                           //Feedback
                           "Mode_HMI_Feedback_Tag(1)" := "Control_DB".LCnv_Control[#i].Mode;
                           "Enabled_HMI_Feedback_Tag(1)" := "Control_DB".LCnv_Control[#i].Enabled;
                           "Error_HMI_Feedback_Tag(1)" := "Control_DB".LCnv_Control[#i].Error;
                           "Warning_HMI_Feedback_Tag(1)" := "Control_DB".LCnv_Control[#i].Warning;
                           "Stopped_HMI_Feedback_Tag(1)" := "Control_DB".LCnv_Control[#i].Stopped;
                           "Running_HMI_Feedback_Tag(1)" := "Control_DB".LCnv_Control[#i].Running;
                           "Ready_For_Task_HMI_Feedback_Tag(1)" := "Control_DB".LCnv_Control[#i].Ready_For_Task;
                           "Cnv_Occupied_HMI_Feedback_Tag(1)" := "Control_DB".LCnv_Control[#i].Cnv_Occupied;
                           "Shuttle_in_place_HMI_Feedback_Tag(1)" := "Control_DB".LCnv_Control[#i].Shuttle_In_Place;
                           "Current_Task_Type_HMI_Feedback_Tag(1)" := "Control_DB".LCnv_Control[#i].Current_Task_Type;
                           "Current_Task_ID_HMI_Feedback_Tag(1)" := "Control_DB".LCnv_Control[#i].Current_Task_ID;
                           "SM_State_HMI_Feedback_Tag(1)" := "Control_DB".LCnv_Control[#i].SM_State;
                           IF "Control_DB".LCnv_Control[#i].Motor.Forward THEN
                               "Motor_Direction_HMI_Feedback_Tag(1)" := 1;
                           ELSIF "Control_DB".LCnv_Control[#i].Motor.Reverse THEN
                               "Motor_Direction_HMI_Feedback_Tag(1)" := 2;
                           ELSE
                               "Motor_Direction_HMI_Feedback_Tag(1)" := 0;
                           END_IF;
                           "Motor_Speed_Requested_HMI_Feedback_Tag(1)" := "Control_DB".LCnv_Control[#i].Motor.Speed;
                           "Motor_Speed_Actual_HMI_Feedback_Tag(1)" := "Control_DB".LCnv_Control[#i].Motor.Speed_Actual;
                           "Transfer_To_ID_HMI_Tag(1)" := "Control_DB".LCnv_Control[#i].Instruction.Transfer_To_ID;
                           "Transfer_From_ID_HMI_Tag(1)" := "Control_DB".LCnv_Control[#i].Instruction.Transfer_From_ID;

                           //Instructions
                           IF "HMI_DB".ScreenNo = 2 THEN
                               "Control_DB".LCnv_Control[#i].Instruction.Stop := "Stop_HMI_Tag(1)";
                               "Control_DB".LCnv_Control[#i].Instruction.Execute := "Manual_Fwd_HMI_Tag(1)" OR "Manual_Bwd_HMI_Tag(1)";
                               "Control_DB".LCnv_Control[#i].Instruction.Mode_Change := "Mode_Change_HMI_Tag(1)";
                               "Control_DB".LCnv_Control[#i].Instruction.Enable := "Enable_HMI_Tag(1)";
                               IF "Control_DB".LCnv_Control[#i].Mode <> 3 THEN
                                   "Control_DB".LCnv_Control[#i].Instruction.Foward := "Manual_Fwd_HMI_Tag(1)";
                                   "Control_DB".LCnv_Control[#i].Instruction.Backward := "Manual_Bwd_HMI_Tag(1)";
                                   "Control_DB".LCnv_Control[#i].Instruction.Start_Transfer := "Start_Transfer_HMI_Tag(1)";
                                   IF "Control_DB".LCnv_Control[#i].Mode = 1 THEN
                                       "Control_DB".LCnv_Control[#i].Instruction.Start_Transfer_Backward := "Transfer_Backward(1)";
                                   END_IF;
                                   "Control_DB".LCnv_Control[#i].Safety_Stop_Cnrl.Instruction.Manual_Extend := "Manual_Sfty_Stopper_Up(1)";
                                   "Control_DB".LCnv_Control[#i].Safety_Stop_Cnrl.Instruction.Manual_Retract := "Manual_Sfty_Stopper_Down(1)";

                                   "Control_DB".LCnv_Control[#i].Instruction.Task_ID := "Task_ID_HMI_Tag(1)";
                                   // "Control_DB".LCnv_Control[#i].Instruction.Transfer_To_ID := "Transfer_To_ID_HMI_Tag(1)";
                                   // "Control_DB".LCnv_Control[#i].Instruction.Transfer_From_ID := "Transfer_From_ID_HMI_Tag(1)";
                                   IF "CNV_In_Out(1)" THEN // 0 = Inbound, 1 = Outbound
                                       "Control_DB".LCnv_Control[#i].Instruction.Transfer_To_ID := DINT#120001 + (#i * 100);
                                       "Control_DB".LCnv_Control[#i].Instruction.Transfer_From_ID := 0;
                                   ELSE
                                       "Control_DB".LCnv_Control[#i].Instruction.Transfer_To_ID := 0;
                                       "Control_DB".LCnv_Control[#i].Instruction.Transfer_From_ID := DINT#120001 + (#i * 100);
                                   END_IF;
                               END_IF;
                           END_IF;
                       END_IF;
                   END_FOR;
               END_REGION

               REGION INBOUND CONVEYOR
                   IF "CNV_ID_HMI_Tag(1)" = "Settings_DB".Inbound_Cnv_Settings.ID THEN
                       //Sensors
                       "HMI_CNV_Pallet Detect 1(1)" := "Control_DB".Inbound_Cnv."Inputs"."Pallet Detect 1";
                       "HMI_CNV_Pallet Detect 2(1)" := "Control_DB".Inbound_Cnv.Inputs."Pallet Detect 2";

                       //Feedback
                       "Mode_HMI_Feedback_Tag(1)" := "Control_DB".Inbound_Cnv.Mode;
                       "Enabled_HMI_Feedback_Tag(1)" := "Control_DB".Inbound_Cnv.Enabled;
                       "Error_HMI_Feedback_Tag(1)" := "Control_DB".Inbound_Cnv.Error;
                       "Warning_HMI_Feedback_Tag(1)" := "Control_DB".Inbound_Cnv.Warning;
                       "Stopped_HMI_Feedback_Tag(1)" := "Control_DB".Inbound_Cnv.Stopped;
                       "Running_HMI_Feedback_Tag(1)" := "Control_DB".Inbound_Cnv.Running;
                       "Ready_For_Task_HMI_Feedback_Tag(1)" := "Control_DB".Inbound_Cnv.Ready_For_Task;
                       "Cnv_Occupied_HMI_Feedback_Tag(1)" := "Control_DB".Inbound_Cnv.Cnv_Occupied;
                       "Current_Task_Type_HMI_Feedback_Tag(1)" := "Control_DB".Inbound_Cnv.Current_Task_Type;
                       "Current_Task_ID_HMI_Feedback_Tag(1)" := "Control_DB".Inbound_Cnv.Current_Task_ID;
                       "SM_State_HMI_Feedback_Tag(1)" := "Control_DB".Inbound_Cnv.SM_State;
                       IF "Control_DB".Inbound_Cnv.Motor.Forward THEN
                           "Motor_Direction_HMI_Feedback_Tag(1)" := 1;
                       ELSIF "Control_DB".Inbound_Cnv.Motor.Reverse THEN
                           "Motor_Direction_HMI_Feedback_Tag(1)" := 2;
                       ELSE
                           "Motor_Direction_HMI_Feedback_Tag(1)" := 0;
                       END_IF;
                       "Motor_Speed_Requested_HMI_Feedback_Tag(1)" := "Control_DB".Inbound_Cnv.Motor.Speed;
                       "Motor_Speed_Actual_HMI_Feedback_Tag(1)" := "Control_DB".Inbound_Cnv.Motor.Speed_Actual;
                       "Transfer_To_ID_HMI_Tag(1)" := "Control_DB".Inbound_Cnv.Instruction.Transfer_To_ID;
                       "Transfer_From_ID_HMI_Tag(1)" := "Control_DB".Inbound_Cnv.Instruction.Transfer_From_ID;

                       //Instructions
                       IF "HMI_DB".ScreenNo = 2 THEN
                           "Control_DB".Inbound_Cnv.Instruction.Stop := "Stop_HMI_Tag(1)";
                           "Control_DB".Inbound_Cnv.Instruction.Execute := "Manual_Fwd_HMI_Tag(1)" OR "Manual_Bwd_HMI_Tag(1)";
                           "Control_DB".Inbound_Cnv.Instruction.Mode_Change := "Mode_Change_HMI_Tag(1)";
                           "Control_DB".Inbound_Cnv.Instruction.Enable := "Enable_HMI_Tag(1)";
                           IF "Control_DB".Inbound_Cnv.Mode <> 3 THEN
                               "Control_DB".Inbound_Cnv.Instruction.Foward := "Manual_Fwd_HMI_Tag(1)";
                               "Control_DB".Inbound_Cnv.Instruction.Backward := "Manual_Bwd_HMI_Tag(1)";
                               "Control_DB".Inbound_Cnv.Instruction.Start_Transfer := "Start_Transfer_HMI_Tag(1)";
                               IF "Control_DB".Inbound_Cnv.Mode = 1 THEN
                                   "Control_DB".Inbound_Cnv.Instruction.Start_Transfer_Backward := "Transfer_Backward(1)";
                               END_IF;
                               "Control_DB".Inbound_Cnv.Instruction.Task_ID := "Task_ID_HMI_Tag(1)";
                               "Control_DB".Inbound_Cnv.Instruction.Transfer_To_ID := "Settings_DB".PopUp_Cnv_Settings[1].ID;
                           END_IF;
                       END_IF;
                   END_IF;
               END_REGION

               REGION OUTBOUND CONVEYOR
                   IF "CNV_ID_HMI_Tag(1)" = "Settings_DB".Outbound_Cnv_Settings.ID THEN
                       //Sensors
                       "HMI_CNV_Pallet Detect 1(1)" := "Control_DB".Outbound_Cnv.Inputs."Pallet Detect";

                       //Feedback
                       "Mode_HMI_Feedback_Tag(1)" := "Control_DB".Outbound_Cnv.Mode;
                       "Enabled_HMI_Feedback_Tag(1)" := "Control_DB".Outbound_Cnv.Enabled;
                       "Error_HMI_Feedback_Tag(1)" := "Control_DB".Outbound_Cnv.Error;
                       "Warning_HMI_Feedback_Tag(1)" := "Control_DB".Outbound_Cnv.Warning;
                       "Stopped_HMI_Feedback_Tag(1)" := "Control_DB".Outbound_Cnv.Stopped;
                       "Running_HMI_Feedback_Tag(1)" := "Control_DB".Outbound_Cnv.Running;
                       "Ready_For_Task_HMI_Feedback_Tag(1)" := "Control_DB".Outbound_Cnv.Ready_For_Task;
                       "Cnv_Occupied_HMI_Feedback_Tag(1)" := "Control_DB".Outbound_Cnv.Cnv_Occupied;
                       "Shuttle_in_place_HMI_Feedback_Tag(1)" := "Control_DB".Outbound_Cnv.Shuttle_In_Place;
                       "Current_Task_Type_HMI_Feedback_Tag(1)" := "Control_DB".Outbound_Cnv.Current_Task_Type;
                       "Current_Task_ID_HMI_Feedback_Tag(1)" := "Control_DB".Outbound_Cnv.Current_Task_ID;
                       "SM_State_HMI_Feedback_Tag(1)" := "Control_DB".Outbound_Cnv.SM_State;
                       IF "Control_DB".Outbound_Cnv.Motor.Forward THEN
                           "Motor_Direction_HMI_Feedback_Tag(1)" := 1;
                       ELSIF "Control_DB".Outbound_Cnv.Motor.Reverse THEN
                           "Motor_Direction_HMI_Feedback_Tag(1)" := 2;
                       ELSE
                           "Motor_Direction_HMI_Feedback_Tag(1)" := 0;
                       END_IF;
                       "Motor_Speed_Requested_HMI_Feedback_Tag(1)" := "Control_DB".Outbound_Cnv.Motor.Speed;
                       "Motor_Speed_Actual_HMI_Feedback_Tag(1)" := "Control_DB".Outbound_Cnv.Motor.Speed_Actual;
                       "Transfer_To_ID_HMI_Tag(1)" := "Control_DB".Outbound_Cnv.Instruction.Transfer_To_ID;
                       "Transfer_From_ID_HMI_Tag(1)" := "Control_DB".Outbound_Cnv.Instruction.Transfer_From_ID;

                       //Instructions
                       IF "HMI_DB".ScreenNo = 2 THEN
                           "Control_DB".Outbound_Cnv.Instruction.Stop := "Stop_HMI_Tag(1)";
                           "Control_DB".Outbound_Cnv.Instruction.Execute := "Manual_Fwd_HMI_Tag(1)" OR "Manual_Bwd_HMI_Tag(1)";
                           "Control_DB".Outbound_Cnv.Instruction.Mode_Change := "Mode_Change_HMI_Tag(1)";
                           "Control_DB".Outbound_Cnv.Instruction.Enable := "Enable_HMI_Tag(1)";
                           IF "Control_DB".Outbound_Cnv.Mode <> 3 THEN
                               "Control_DB".Outbound_Cnv.Instruction.Foward := "Manual_Fwd_HMI_Tag(1)";
                               "Control_DB".Outbound_Cnv.Instruction.Backward := "Manual_Bwd_HMI_Tag(1)";
                               "Control_DB".Outbound_Cnv.Instruction.Start_Transfer := "Start_Transfer_HMI_Tag(1)";
                               IF "Control_DB".Outbound_Cnv.Mode = 1 THEN
                                   "Control_DB".Outbound_Cnv.Instruction.Start_Transfer_Backward := "Transfer_Backward(1)";
                               END_IF;
                               "Control_DB".Outbound_Cnv.Instruction.Task_ID := "Task_ID_HMI_Tag(1)";
                               "Control_DB".Outbound_Cnv.Instruction.Transfer_From_ID := "Settings_DB".PopUp_Cnv_Settings[4].ID;
                           END_IF;
                       END_IF;
                   END_IF;
               END_REGION

               REGION POPUP CONVEYORS
                   IF "CNV_ID_HMI_Tag(1)" = "Settings_DB".PopUp_Cnv_Settings[1].ID THEN
                       "HMI_CNV_Pallet Detect 1(1)" := "PopUp Conveyor 1 - Pallet sensor";
                       "HMI_CNV_Pallet Detect 2(1)" := "Pick Station";
                   ELSIF "CNV_ID_HMI_Tag(1)" = "Settings_DB".PopUp_Cnv_Settings[2].ID THEN
                       "HMI_CNV_Pallet Detect 1(1)" := "PopUp Conveyor 2 - Pallet Present 1";
                       "HMI_CNV_Pallet Detect 2(1)" := "PopUp Conveyor 2 - Pallet present 2";
                       "HMI_CNV_Pallet Detect 3(1)" := "PopUp Conveyor 2 - Pallet present 3";
                       "HMI_CNV_Pallet Detect 4(1)" := "PopUp Conveyor 2 - Pallet present 4";
                       "HMI_CNV_Pallet Detect 5(1)" := "PopUp Conveyor 2 - Pallet present 5";
                   ELSIF "CNV_ID_HMI_Tag(1)" = "Settings_DB".PopUp_Cnv_Settings[3].ID THEN
                       "HMI_CNV_Pallet Detect 1(1)" := "PopUp Conveyor 3 - Pallet present 1";
                   ELSIF "CNV_ID_HMI_Tag(1)" = "Settings_DB".PopUp_Cnv_Settings[4].ID THEN
                       "HMI_CNV_Pallet Detect 1(1)" := "PopUp Conveyor 4 - Pallet present 1";
                       "HMI_CNV_Pallet Detect 2(1)" := "Pick Station";
                   END_IF;

                   FOR #i := 1 TO 4 DO
                       IF "CNV_ID_HMI_Tag(1)" = "Settings_DB".PopUp_Cnv_Settings[#i].ID THEN
                           //Sensors
                           IF "Control_DB".PopUp_Cnv[#i].Inputs."Lift Up" AND NOT "Control_DB".PopUp_Cnv[#i].Inputs."Lift Down" THEN
                               "UP_DOWN(1)" := 1;
                           ELSIF NOT "Control_DB".PopUp_Cnv[#i].Inputs."Lift Up" AND "Control_DB".PopUp_Cnv[#i].Inputs."Lift Down" THEN
                               "UP_DOWN(1)" := 2;
                           ELSE
                               "UP_DOWN(1)" := 0;
                           END_IF;
                           IF "CNV_ID_HMI_Tag(1)" = "Settings_DB".PopUp_Cnv_Settings[#i].ID THEN
                               //Feedback
                               "Mode_HMI_Feedback_Tag(1)" := "Control_DB".PopUp_Cnv[#i].Mode;
                               "Enabled_HMI_Feedback_Tag(1)" := "Control_DB".PopUp_Cnv[#i].Enabled;
                               "Error_HMI_Feedback_Tag(1)" := "Control_DB".PopUp_Cnv[#i].Error;
                               "Warning_HMI_Feedback_Tag(1)" := "Control_DB".PopUp_Cnv[#i].Warning;
                               "Stopped_HMI_Feedback_Tag(1)" := "Control_DB".PopUp_Cnv[#i].Stopped;
                               "Running_HMI_Feedback_Tag(1)" := "Control_DB".PopUp_Cnv[#i].Running;
                               "Ready_For_Task_HMI_Feedback_Tag(1)" := "Control_DB".PopUp_Cnv[#i].Ready_For_Task;
                               "Cnv_Occupied_HMI_Feedback_Tag(1)" := "Control_DB".PopUp_Cnv[#i].Cnv_Occupied;
                               "Current_Task_Type_HMI_Feedback_Tag(1)" := "Control_DB".PopUp_Cnv[#i].Current_Task_Type;
                               "Current_Task_ID_HMI_Feedback_Tag(1)" := "Control_DB".PopUp_Cnv[#i].Current_Task_ID;
                               "SM_State_HMI_Feedback_Tag(1)" := "Control_DB".PopUp_Cnv[#i].SM_State;
                               "Transfer_To_ID_HMI_Tag(1)" := "Control_DB".PopUp_Cnv[#i].Instruction.Transfer_To_ID;
                               "Transfer_From_ID_HMI_Tag(1)" := "Control_DB".PopUp_Cnv[#i].Instruction.Transfer_From_ID;
                               IF "Control_DB".PopUp_Cnv[#i].Roller_Motor.Status.%X0 THEN
                                   IF "Control_DB".PopUp_Cnv[#i].Roller_Motor.Forward THEN
                                       "Motor_Direction_HMI_Feedback_Tag(1)" := 1;
                                   ELSIF "Control_DB".PopUp_Cnv[#i].Roller_Motor.Reverse THEN
                                       "Motor_Direction_HMI_Feedback_Tag(1)" := 2;
                                   ELSE
                                       "Motor_Direction_HMI_Feedback_Tag(1)" := 0;
                                   END_IF;
                                   "Motor_Speed_Requested_HMI_Feedback_Tag(1)" := REAL_TO_UINT("Control_DB".PopUp_Cnv[#i].Roller_Motor.Speed);
                                   "Motor_Speed_Actual_HMI_Feedback_Tag(1)" := REAL_TO_UINT("Control_DB".PopUp_Cnv[#i].Roller_Motor.Speed_Actual);
                               ELSIF "Control_DB".PopUp_Cnv[#i].Chain_Motor.Status.%X0 = 1 THEN
                                   IF "Control_DB".PopUp_Cnv[#i].Chain_Motor.Forward THEN
                                       "Motor_Direction_HMI_Feedback_Tag(1)" := 1;
                                   ELSIF "Control_DB".PopUp_Cnv[#i].Chain_Motor.Reverse THEN
                                       "Motor_Direction_HMI_Feedback_Tag(1)" := 2;
                                   ELSE
                                       "Motor_Direction_HMI_Feedback_Tag(1)" := 0;
                                   END_IF;
                                   "Motor_Speed_Requested_HMI_Feedback_Tag(1)" := REAL_TO_UINT("Control_DB".PopUp_Cnv[#i].Chain_Motor.Speed);
                                   "Motor_Speed_Actual_HMI_Feedback_Tag(1)" := REAL_TO_UINT("Control_DB".PopUp_Cnv[#i].Chain_Motor.Speed_Actual);
                               ELSIF "Control_DB".PopUp_Cnv[#i].Lift_Motor.Status.%X0 = 1 THEN
                                   IF "Control_DB".PopUp_Cnv[#i].Lift_Motor.Forward THEN
                                       "Motor_Direction_HMI_Feedback_Tag(1)" := 1;
                                   ELSIF "Control_DB".PopUp_Cnv[#i].Lift_Motor.Reverse THEN
                                       "Motor_Direction_HMI_Feedback_Tag(1)" := 2;
                                   ELSE
                                       "Motor_Direction_HMI_Feedback_Tag(1)" := 0;
                                   END_IF;
                                   "Motor_Speed_Requested_HMI_Feedback_Tag(1)" := REAL_TO_UINT("Control_DB".PopUp_Cnv[#i].Lift_Motor.Speed);
                                   "Motor_Speed_Actual_HMI_Feedback_Tag(1)" := REAL_TO_UINT("Control_DB".PopUp_Cnv[#i].Lift_Motor.Speed_Actual);
                               END_IF;

                               //Instructions
                               IF "HMI_DB".ScreenNo = 2 THEN
                                   "Control_DB".PopUp_Cnv[#i].Instruction.Stop := "Stop_HMI_Tag(1)";
                                   "Control_DB".PopUp_Cnv[#i].Instruction.Execute := "Manual_Fwd_HMI_Tag(1)" OR "Manual_Bwd_HMI_Tag(1)";
                                   "Control_DB".PopUp_Cnv[#i].Instruction.Mode_Change := "Mode_Change_HMI_Tag(1)";
                                   "Control_DB".PopUp_Cnv[#i].Instruction.Enable := "Enable_HMI_Tag(1)";
                                   IF "Control_DB".PopUp_Cnv[#i].Mode <> 3 THEN
                                       IF "Control_DB".PopUp_Cnv[#i].Inputs."Lift Up" THEN
                                           "Control_DB".PopUp_Cnv[#i].Instruction.Roller_Fwd := "Manual_Fwd_HMI_Tag(1)";
                                           "Control_DB".PopUp_Cnv[#i].Instruction.Roller_Bwd := "Manual_Bwd_HMI_Tag(1)";
                                       ELSIF "Control_DB".PopUp_Cnv[#i].Inputs."Lift Down" THEN
                                           "Control_DB".PopUp_Cnv[#i].Instruction.Chain_Fwd := "Manual_Fwd_HMI_Tag(1)";
                                           "Control_DB".PopUp_Cnv[#i].Instruction.Chain_Bwd := "Manual_Bwd_HMI_Tag(1)";
                                       END_IF;
                                       "Control_DB".PopUp_Cnv[#i].Instruction.Start_Transfer := "Start_Transfer_HMI_Tag(1)";
                                       IF "Control_DB".PopUp_Cnv[#i].Mode = 1 THEN
                                           "Control_DB".PopUp_Cnv[#i].Instruction.Start_Transfer_Backward := "Transfer_Backward(1)";
                                       END_IF;
                                       "Control_DB".PopUp_Cnv[#i].Instruction.Lift_Up := "Manual_Sfty_Stopper_Up(1)";
                                       "Control_DB".PopUp_Cnv[#i].Instruction.Lift_Down := "Manual_Sfty_Stopper_Down(1)";
                                       "Control_DB".PopUp_Cnv[#i].Instruction.Task_ID := "Task_ID_HMI_Tag(1)";
                                       CASE #i OF
                                           1:
                                               IF "CNV_In_Out(1)" AND "Control_DB".PopUp_Cnv[1].Inputs."Lift Up" THEN // 0 = Inbound, 1 = Outbound
                                                   "Control_DB".PopUp_Cnv[#i].Instruction.Transfer_To_ID := "Settings_DB".PopUp_Cnv_Settings[2].ID;
                                                   "Control_DB".PopUp_Cnv[#i].Instruction.Transfer_From_ID := 0;
                                               ELSIF NOT "CNV_In_Out(1)" AND "Control_DB".PopUp_Cnv[1].Inputs."Lift Down" AND "Pick Station" THEN // 0 = Inbound, 1 = Outbound
                                                   "Control_DB".PopUp_Cnv[#i].Instruction.Transfer_To_ID := 0;
                                                   "Control_DB".PopUp_Cnv[#i].Instruction.Transfer_From_ID := "Settings_DB".Pick_Cnv_Settings.ID;
                                               ELSIF NOT "CNV_In_Out(1)" AND "Control_DB".PopUp_Cnv[1].Inputs."Lift Up" THEN // 0 = Inbound, 1 = Outbound
                                                   "Control_DB".PopUp_Cnv[#i].Instruction.Transfer_To_ID := 0;
                                                   "Control_DB".PopUp_Cnv[#i].Instruction.Transfer_From_ID := "Settings_DB".Inbound_Cnv_Settings.ID;
                                               ELSE
                                                   "Control_DB".PopUp_Cnv[#i].Instruction.Transfer_To_ID := 0;
                                                   "Control_DB".PopUp_Cnv[#i].Instruction.Transfer_From_ID := 0;
                                               END_IF;

                                           2:
                                               IF NOT "CNV_In_Out(1)" AND "Control_DB".PopUp_Cnv[2].Inputs."Lift Up" THEN // UP
                                                   "Control_DB".PopUp_Cnv[#i].Instruction.Transfer_To_ID := 0;
                                                   "Control_DB".PopUp_Cnv[#i].Instruction.Transfer_From_ID := "Settings_DB".PopUp_Cnv_Settings[1].ID;
                                               ELSIF NOT "CNV_In_Out(1)" AND "Control_DB".PopUp_Cnv[2].Inputs."Lift Down" THEN //DOWN
                                                   "Control_DB".PopUp_Cnv[#i].Instruction.Transfer_To_ID := 0;
                                                   "Control_DB".PopUp_Cnv[#i].Instruction.Transfer_From_ID := "Settings_DB".ECnv_Settings.ID;
                                               ELSIF "CNV_In_Out(1)" AND "Control_DB".PopUp_Cnv[2].Inputs."Lift Down" AND NOT "VTD_POPUP2(1)" THEN //DOWN
                                                   "Control_DB".PopUp_Cnv[#i].Instruction.Transfer_To_ID := "Settings_DB".ECnv_Settings.ID;
                                                   "Control_DB".PopUp_Cnv[#i].Instruction.Transfer_From_ID := 0;
                                               ELSIF "CNV_In_Out(1)" AND "Control_DB".PopUp_Cnv[2].Inputs."Lift Down" AND "VTD_POPUP2(1)" THEN //DOWN
                                                   "Control_DB".PopUp_Cnv[#i].Instruction.Transfer_To_ID := "Settings_DB".PopUp_Cnv_Settings[3].ID;
                                                   "Control_DB".PopUp_Cnv[#i].Instruction.Transfer_From_ID := 0;
                                               ELSE
                                                   "Control_DB".PopUp_Cnv[#i].Instruction.Transfer_To_ID := 0;
                                                   "Control_DB".PopUp_Cnv[#i].Instruction.Transfer_From_ID := 0;
                                               END_IF;

                                           3:
                                               IF NOT "CNV_In_Out(1)" AND "Control_DB".PopUp_Cnv[3].Inputs."Lift Down" THEN //inbound chain
                                                   "Control_DB".PopUp_Cnv[#i].Instruction.Transfer_To_ID := 0;
                                                   "Control_DB".PopUp_Cnv[#i].Instruction.Transfer_From_ID := "Settings_DB".PopUp_Cnv_Settings[2].ID;
                                               ELSIF "CNV_In_Out(1)" AND "Control_DB".PopUp_Cnv[3].Inputs."Lift Up" THEN //DOWN
                                                   "Control_DB".PopUp_Cnv[#i].Instruction.Transfer_To_ID := "Settings_DB".PopUp_Cnv_Settings[4].ID;
                                                   "Control_DB".PopUp_Cnv[#i].Instruction.Transfer_From_ID := 0;
                                               ELSE
                                                   "Control_DB".PopUp_Cnv[#i].Instruction.Transfer_To_ID := 0;
                                                   "Control_DB".PopUp_Cnv[#i].Instruction.Transfer_From_ID := 0;
                                               END_IF;

                                           4:
                                               IF "CNV_In_Out(1)" AND "Control_DB".PopUp_Cnv[4].Inputs."Lift Up" THEN // 0 = Inbound, 1 = Outbound
                                                   "Control_DB".PopUp_Cnv[#i].Instruction.Transfer_To_ID := "Settings_DB".Outbound_Cnv_Settings.ID;
                                                   "Control_DB".PopUp_Cnv[#i].Instruction.Transfer_From_ID := 0;
                                               ELSIF "CNV_In_Out(1)" AND "Control_DB".PopUp_Cnv[4].Inputs."Lift Down" AND "Pick Station" THEN // 0 = Inbound, 1 = Outbound
                                                   "Control_DB".PopUp_Cnv[#i].Instruction.Transfer_To_ID := "Settings_DB".Pick_Cnv_Settings.ID;
                                                   "Control_DB".PopUp_Cnv[#i].Instruction.Transfer_From_ID := 0;
                                               ELSIF NOT "CNV_In_Out(1)" AND "Control_DB".PopUp_Cnv[4].Inputs."Lift Up" THEN // 0 = Inbound, 1 = Outbound
                                                   "Control_DB".PopUp_Cnv[#i].Instruction.Transfer_To_ID := 0;
                                                   "Control_DB".PopUp_Cnv[#i].Instruction.Transfer_From_ID := "Settings_DB".PopUp_Cnv_Settings[3].ID;
                                               ELSE
                                                   "Control_DB".PopUp_Cnv[#i].Instruction.Transfer_To_ID := 0;
                                                   "Control_DB".PopUp_Cnv[#i].Instruction.Transfer_From_ID := 0;
                                               END_IF;
                                       END_CASE;
                                   END_IF;
                               END_IF;
                           END_IF;
                       END_IF;
                   END_FOR;
               END_REGION

               REGION PICK CONVEYOR
                   IF "CNV_ID_HMI_Tag(1)" = "Settings_DB".Pick_Cnv_Settings.ID THEN
                       //Sensors
                       "HMI_CNV_Pallet Detect 1(1)" := "Control_DB".Pick_Station.Cnv_Occupied;

                       //Feedback
                       "Mode_HMI_Feedback_Tag(1)" := "Control_DB".Pick_Station.Mode;
                       "Enabled_HMI_Feedback_Tag(1)" := "Control_DB".Pick_Station.Enabled;
                       "Error_HMI_Feedback_Tag(1)" := "Control_DB".Pick_Station.Error;
                       "Warning_HMI_Feedback_Tag(1)" := "Control_DB".Pick_Station.Warning;
                       "Stopped_HMI_Feedback_Tag(1)" := "Control_DB".Pick_Station.Stopped;
                       "Running_HMI_Feedback_Tag(1)" := "Control_DB".Pick_Station.Running;
                       "Ready_For_Task_HMI_Feedback_Tag(1)" := "Control_DB".Pick_Station.Ready_For_Task;
                       "Cnv_Occupied_HMI_Feedback_Tag(1)" := "Control_DB".Pick_Station.Cnv_Occupied;
                       // "Shuttle_in_place_HMI_Feedback_Tag(1)" := "Control_DB".Pick_Station.Shuttle_In_Place;
                       "Current_Task_Type_HMI_Feedback_Tag(1)" := "Control_DB".Pick_Station.Current_Task_Type;
                       "Current_Task_ID_HMI_Feedback_Tag(1)" := "Control_DB".Pick_Station.Current_Task_ID;
                       "SM_State_HMI_Feedback_Tag(1)" := "Control_DB".Pick_Station.SM_State;
                       IF "Control_DB".Pick_Station.Motor.Forward THEN
                           "Motor_Direction_HMI_Feedback_Tag(1)" := 1;
                       ELSIF "Control_DB".Pick_Station.Motor.Reverse THEN
                           "Motor_Direction_HMI_Feedback_Tag(1)" := 2;
                       ELSE
                           "Motor_Direction_HMI_Feedback_Tag(1)" := 0;
                       END_IF;
                       "Motor_Speed_Requested_HMI_Feedback_Tag(1)" := "Control_DB".Pick_Station.Motor.Speed;
                       "Motor_Speed_Actual_HMI_Feedback_Tag(1)" := "Control_DB".Pick_Station.Motor.Speed_Actual;
                       "Transfer_To_ID_HMI_Tag(1)" := "Control_DB".Pick_Station.Instruction.Transfer_To_ID;
                       "Transfer_From_ID_HMI_Tag(1)" := "Control_DB".Pick_Station.Instruction.Transfer_From_ID;

                       //Instructions
                       IF "HMI_DB".ScreenNo = 2 THEN
                           "Control_DB".Pick_Station.Instruction.Stop := "Stop_HMI_Tag(1)";
                           "Control_DB".Pick_Station.Instruction.Execute := "Manual_Fwd_HMI_Tag(1)" OR "Manual_Bwd_HMI_Tag(1)";
                           "Control_DB".Pick_Station.Instruction.Mode_Change := "Mode_Change_HMI_Tag(1)";
                           "Control_DB".Pick_Station.Instruction.Enable := "Enable_HMI_Tag(1)";
                           IF "Control_DB".Pick_Station.Mode <> 3 THEN
                               "Control_DB".Pick_Station.Instruction.Foward := "Manual_Fwd_HMI_Tag(1)";
                               "Control_DB".Pick_Station.Instruction.Backward := "Manual_Bwd_HMI_Tag(1)";
                               "Control_DB".Pick_Station.Instruction.Start_Transfer := "Start_Transfer_HMI_Tag(1)";
                               IF "Control_DB".Pick_Station.Mode = 1 THEN
                                   "Control_DB".Pick_Station.Instruction.Start_Transfer_Backward := "Transfer_Backward(1)";
                               END_IF;
                               "Control_DB".Pick_Station.Instruction.Task_ID := "Task_ID_HMI_Tag(1)";
                               "Control_DB".Pick_Station.Instruction.Transfer_From_ID := "Settings_DB".PopUp_Cnv_Settings[4].ID;
                               "Control_DB".Pick_Station.Instruction.Transfer_To_ID := "Settings_DB".PopUp_Cnv_Settings[1].ID;
                           END_IF;
                       END_IF;
                   END_IF;
               END_REGION
           END_IF;
       END_REGION
   END_REGION

   "IEC_Timer_0_DB_4".TON(IN := "Screen_DB".Charge_VTD OR "Screen_DB".Charge_Cnv OR "Screen_DB".Charge_VTD_Commands OR "Screen_DB".Charge_Cnv_Commands,
                          PT := T#1S);

   IF "IEC_Timer_0_DB_4".Q THEN
       "Screen_DB".Charge_VTD := FALSE;
       "Screen_DB".Charge_Cnv := FALSE;
       "Screen_DB".Charge_VTD_Commands := FALSE;
       "Screen_DB".Charge_Cnv_Commands := FALSE;
   END_IF;

   "Control_DB".ECnv_Control.Instruction.Reset := "Reset_HMI_Tag" OR "Reset_All" OR "Reset_HMI_Tag(1)";
   "Control_DB".LCnv_Control[1].Instruction.Reset := "Reset_HMI_Tag" OR "Reset_HMI_Tag(1)" OR "Reset_All";
   "Control_DB".LCnv_Control[1].Instruction.Reset := "Reset_HMI_Tag" OR "Reset_HMI_Tag(1)" OR "Reset_All";
   "Control_DB".LCnv_Control[2].Instruction.Reset := "Reset_HMI_Tag" OR "Reset_HMI_Tag(1)" OR "Reset_All";
   "Control_DB".LCnv_Control[2].Instruction.Reset := "Reset_HMI_Tag" OR "Reset_HMI_Tag(1)" OR "Reset_All";
   "Control_DB".LCnv_Control[3].Instruction.Reset := "Reset_HMI_Tag" OR "Reset_HMI_Tag(1)" OR "Reset_All";
   "Control_DB".LCnv_Control[3].Instruction.Reset := "Reset_HMI_Tag" OR "Reset_HMI_Tag(1)" OR "Reset_All";
   "Control_DB".Inbound_Cnv.Instruction.Reset := "Reset_HMI_Tag" OR "Reset_HMI_Tag(1)" OR "Reset_All";
   "Control_DB".Outbound_Cnv.Instruction.Reset := "Reset_HMI_Tag" OR "Reset_HMI_Tag(1)" OR "Reset_All";
   "Control_DB".Pick_Station.Instruction.Reset := "Reset_HMI_Tag" OR "Reset_HMI_Tag(1)" OR "Reset_All";
   "Control_DB".Pick_Station.Instruction.Reset := "Reset_HMI_Tag" OR "Reset_HMI_Tag(1)" OR "Reset_All";
   "Control_DB".PopUp_Cnv[1].Instruction.Reset := "Reset_HMI_Tag" OR "Reset_HMI_Tag(1)" OR "Reset_All";
   "Control_DB".PopUp_Cnv[2].Instruction.Reset := "Reset_HMI_Tag" OR "Reset_HMI_Tag(1)" OR "Reset_All";
   "Control_DB".PopUp_Cnv[3].Instruction.Reset := "Reset_HMI_Tag" OR "Reset_HMI_Tag(1)" OR "Reset_All";
   "Control_DB".PopUp_Cnv[4].Instruction.Reset := "Reset_HMI_Tag" OR "Reset_HMI_Tag(1)" OR "Reset_All";


   //START TRANSFER BACKWARD VISIBILITY
   IF "Mode_Change_HMI_Tag" = 1 AND "Mode_Change_HMI_Tag(1)" = 1 THEN
       "Transfer_Backward_Visibility" :=
       //inbound - popup 1
       ("CNV_ID_HMI_Tag" = "Settings_DB".Inbound_Cnv_Settings.ID AND "CNV_ID_HMI_Tag(1)" = "Settings_DB".PopUp_Cnv_Settings[1].ID) OR
       ("CNV_ID_HMI_Tag" = "Settings_DB".PopUp_Cnv_Settings[1].ID AND "CNV_ID_HMI_Tag(1)" = "Settings_DB".Inbound_Cnv_Settings.ID) OR
       //POPUP1 - popup 2
       ("CNV_ID_HMI_Tag" = "Settings_DB".PopUp_Cnv_Settings[1].ID AND "CNV_ID_HMI_Tag(1)" = "Settings_DB".PopUp_Cnv_Settings[2].ID) OR
       ("CNV_ID_HMI_Tag" = "Settings_DB".PopUp_Cnv_Settings[2].ID AND "CNV_ID_HMI_Tag(1)" = "Settings_DB".PopUp_Cnv_Settings[1].ID) OR
       //POPUP2 - popup 3
       ("CNV_ID_HMI_Tag" = "Settings_DB".PopUp_Cnv_Settings[2].ID AND "CNV_ID_HMI_Tag(1)" = "Settings_DB".PopUp_Cnv_Settings[3].ID) OR
       ("CNV_ID_HMI_Tag" = "Settings_DB".PopUp_Cnv_Settings[3].ID AND "CNV_ID_HMI_Tag(1)" = "Settings_DB".PopUp_Cnv_Settings[2].ID) OR
       //POPUP3 - popup 4
       ("CNV_ID_HMI_Tag" = "Settings_DB".PopUp_Cnv_Settings[3].ID AND "CNV_ID_HMI_Tag(1)" = "Settings_DB".PopUp_Cnv_Settings[4].ID) OR
       ("CNV_ID_HMI_Tag" = "Settings_DB".PopUp_Cnv_Settings[4].ID AND "CNV_ID_HMI_Tag(1)" = "Settings_DB".PopUp_Cnv_Settings[3].ID) OR
       //POPUP4 - POPUP 1
       ("CNV_ID_HMI_Tag" = "Settings_DB".PopUp_Cnv_Settings[4].ID AND "CNV_ID_HMI_Tag(1)" = "Settings_DB".PopUp_Cnv_Settings[1].ID) OR
       ("CNV_ID_HMI_Tag" = "Settings_DB".PopUp_Cnv_Settings[1].ID AND "CNV_ID_HMI_Tag(1)" = "Settings_DB".PopUp_Cnv_Settings[4].ID) OR
       //POPUP4 - OUTBOUND
       ("CNV_ID_HMI_Tag" = "Settings_DB".PopUp_Cnv_Settings[4].ID AND "CNV_ID_HMI_Tag(1)" = "Settings_DB".Outbound_Cnv_Settings.ID) OR
       ("CNV_ID_HMI_Tag" = "Settings_DB".Outbound_Cnv_Settings.ID AND "CNV_ID_HMI_Tag(1)" = "Settings_DB".PopUp_Cnv_Settings[4].ID) OR
       //POPUP2 - EConveyor
       ("CNV_ID_HMI_Tag" = "Settings_DB".PopUp_Cnv_Settings[2].ID AND "CNV_ID_HMI_Tag(1)" = "Settings_DB".ECnv_Settings.ID) OR
       ("CNV_ID_HMI_Tag" = "Settings_DB".ECnv_Settings.ID AND "CNV_ID_HMI_Tag(1)" = "Settings_DB".PopUp_Cnv_Settings[2].ID) OR
       //EConveyor - Buffer 1
       ("CNV_ID_HMI_Tag" = "Settings_DB".ECnv_Settings.ID AND "CNV_ID_HMI_Tag(1)" = "Settings_DB".LCnv_Settings[1].ID) OR
       ("CNV_ID_HMI_Tag" = "Settings_DB".LCnv_Settings[1].ID AND "CNV_ID_HMI_Tag(1)" = "Settings_DB".ECnv_Settings.ID) OR
       //EConveyor - Buffer 2
       ("CNV_ID_HMI_Tag" = "Settings_DB".ECnv_Settings.ID AND "CNV_ID_HMI_Tag(1)" = "Settings_DB".LCnv_Settings[2].ID) OR
       ("CNV_ID_HMI_Tag" = "Settings_DB".LCnv_Settings[2].ID AND "CNV_ID_HMI_Tag(1)" = "Settings_DB".ECnv_Settings.ID) OR
       //EConveyor - Buffer 3
       ("CNV_ID_HMI_Tag" = "Settings_DB".ECnv_Settings.ID AND "CNV_ID_HMI_Tag(1)" = "Settings_DB".LCnv_Settings[3].ID) OR
       ("CNV_ID_HMI_Tag" = "Settings_DB".LCnv_Settings[3].ID AND "CNV_ID_HMI_Tag(1)" = "Settings_DB".ECnv_Settings.ID) OR
       //PICK - POPUP4
       ("CNV_ID_HMI_Tag" = "Settings_DB".Pick_Cnv_Settings.ID AND "CNV_ID_HMI_Tag(1)" = "Settings_DB".PopUp_Cnv_Settings[4].ID) OR
       ("CNV_ID_HMI_Tag" = "Settings_DB".PopUp_Cnv_Settings[4].ID AND "CNV_ID_HMI_Tag(1)" = "Settings_DB".Pick_Cnv_Settings.ID);
   ELSE
       "Transfer_Backward_Visibility" := FALSE;
   END_IF;
END_FUNCTION_BLOCK

FUNCTION "PopUp_Screens" : Void   // FC9, SCL
{ S7_Optimized_Access := 'TRUE' }
VERSION : 0.1
// stored: AutoNumber true, IsIECCheckEnabled false, SetENOAutomatically false, UDAEnableTagReadback false
BEGIN
   //CHARGE SETTINGS CHANGING CONVEYORS SELECTION
   IF "PopUps_DB".Cnv_Select <> "PopUps_DB".Cnv_Select_Old THEN
       "Screen_DB".Charge_Cnv := TRUE;
       "PopUps_DB".Cnv_Select_Old := "PopUps_DB".Cnv_Select;
   END_IF;

   //CHARGE VTD SETTINGS FROM DB
   "R_TRIG_DB"(CLK := "Screen_DB".Charge_VTD);
   IF "R_TRIG_DB".Q THEN
       //VTD SETTINGS
       "PopUps_DB".VTD_Settings := "Settings_DB".VTD_Settings;
       "PopUps_DB".Shuttle_MQTT_Settings := "Settings_DB".Shuttle_MQTT_Settings;
       "Screen_DB".Charge_VTD := 0;
   END_IF;

   //CHARGE CNV SETTINGS FROM DB
   "R_TRIG_DB_4"(CLK := "Screen_DB".Charge_Cnv);
   IF "R_TRIG_DB_4".Q THEN
       "EConveyor_Visibility" := "PConveyor_Visibility" := "IConveyor_Visibility" := "OConveyor_Visibility" := "BConveyor_Visibility" := FALSE;
       //CONVEYORS SETTINGS
       CASE "PopUps_DB".Cnv_Select OF
           120001:
               "PopUps_DB".ECnv_Settings := "Settings_DB".ECnv_Settings;
           100101:
               "PopUps_DB".Buffer_Cnv_Settings := "Settings_DB".LCnv_Settings[1];
           100201:
               "PopUps_DB".Buffer_Cnv_Settings := "Settings_DB".LCnv_Settings[2];
           100301:
               "PopUps_DB".Buffer_Cnv_Settings := "Settings_DB".LCnv_Settings[3];
           130001:
               "PopUps_DB".Inbound_Cnv_Settings := "Settings_DB".Inbound_Cnv_Settings;
           140001:
               "PopUps_DB".Outbound_Cnv_Settings := "Settings_DB".Outbound_Cnv_Settings;
           150001:
               "PopUps_DB".PopUp_Cnv_settings := "Settings_DB".PopUp_Cnv_Settings[1];
           160001:
               "PopUps_DB".PopUp_Cnv_settings := "Settings_DB".PopUp_Cnv_Settings[2];
           170001:
               "PopUps_DB".PopUp_Cnv_settings := "Settings_DB".PopUp_Cnv_Settings[3];
           180001:
               "PopUps_DB".PopUp_Cnv_settings := "Settings_DB".PopUp_Cnv_Settings[4];
           410001:
               "PopUps_DB".Outbound_Cnv_Settings := "Settings_DB".Pick_Cnv_Settings;
       END_CASE;
       // "Screen_DB".Charge_Cnv := 0;
   END_IF;

   //CHARGE VTD SETTINGS FROM HMI
   IF NOT "Screen_DB".Charge_VTD THEN

       IF "HMI_DB".ScreenNo = 7 OR "HMI_DB".ScreenNo = 11 THEN
           "Settings_DB".VTD_Settings := "PopUps_DB".VTD_Settings;
       END_IF;

       //SHUTTLE MQTT SETTINGS
       "Settings_DB".Shuttle_MQTT_Settings := "PopUps_DB".Shuttle_MQTT_Settings;
   END_IF;

   //CHARGE CNV SETTINGS FROM HMI
   IF NOT "Screen_DB".Charge_Cnv THEN
       //CONVEYORS SETTINGS
       IF "HMI_DB".ScreenNo = 8 OR "HMI_DB".ScreenNo = 10 THEN
           CASE "PopUps_DB".Cnv_Select OF
               120001:
                   "Settings_DB".ECnv_Settings := "PopUps_DB".ECnv_Settings;
                   "PConveyor_Visibility" := "IConveyor_Visibility" := "OConveyor_Visibility" := "BConveyor_Visibility" := FALSE;
                   "EConveyor_Visibility" := TRUE;

               100101:
                   "Settings_DB".LCnv_Settings[1] := "PopUps_DB".Buffer_Cnv_Settings;
                   "PConveyor_Visibility" := "IConveyor_Visibility" := "OConveyor_Visibility" := "EConveyor_Visibility" := FALSE;
                   "BConveyor_Visibility" := TRUE;

               100201:
                   "Settings_DB".LCnv_Settings[2] := "PopUps_DB".Buffer_Cnv_Settings;
                   "PConveyor_Visibility" := "IConveyor_Visibility" := "OConveyor_Visibility" := "EConveyor_Visibility" := FALSE;
                   "BConveyor_Visibility" := TRUE;

               100301:
                   "Settings_DB".LCnv_Settings[3] := "PopUps_DB".Buffer_Cnv_Settings;
                   "PConveyor_Visibility" := "IConveyor_Visibility" := "OConveyor_Visibility" := "EConveyor_Visibility" := FALSE;
                   "BConveyor_Visibility" := TRUE;

               130001:
                   "Settings_DB".Inbound_Cnv_Settings := "PopUps_DB".Inbound_Cnv_Settings;
                   "PConveyor_Visibility" := "BConveyor_Visibility" := "OConveyor_Visibility" := "EConveyor_Visibility" := FALSE;
                   "IConveyor_Visibility" := TRUE;

               140001:
                   "Settings_DB".Outbound_Cnv_Settings := "PopUps_DB".Outbound_Cnv_Settings;
                   "PConveyor_Visibility" := "BConveyor_Visibility" := "IConveyor_Visibility" := "EConveyor_Visibility" := FALSE;
                   "OConveyor_Visibility" := TRUE;

               150001:
                   "Settings_DB".PopUp_Cnv_Settings[1] := "PopUps_DB".PopUp_Cnv_settings;
                   "BConveyor_Visibility" := "IConveyor_Visibility" := "OConveyor_Visibility" := "EConveyor_Visibility" := FALSE;
                   "PConveyor_Visibility" := TRUE;

               160001:
                   "Settings_DB".PopUp_Cnv_Settings[2] := "PopUps_DB".PopUp_Cnv_settings;
                   "BConveyor_Visibility" := "IConveyor_Visibility" := "OConveyor_Visibility" := "EConveyor_Visibility" := FALSE;
                   "PConveyor_Visibility" := TRUE;

               170001:
                   "Settings_DB".PopUp_Cnv_Settings[3] := "PopUps_DB".PopUp_Cnv_settings;
                   "BConveyor_Visibility" := "IConveyor_Visibility" := "OConveyor_Visibility" := "EConveyor_Visibility" := FALSE;
                   "PConveyor_Visibility" := TRUE;

               180001:
                   "Settings_DB".PopUp_Cnv_Settings[4] := "PopUps_DB".PopUp_Cnv_settings;
                   "BConveyor_Visibility" := "IConveyor_Visibility" := "OConveyor_Visibility" := "EConveyor_Visibility" := FALSE;
                   "PConveyor_Visibility" := TRUE;

               410001:
                   "Settings_DB".Pick_Cnv_Settings := "PopUps_DB".Outbound_Cnv_Settings;
                   "PConveyor_Visibility" := "BConveyor_Visibility" := "IConveyor_Visibility" := "EConveyor_Visibility" := FALSE;
                   "OConveyor_Visibility" := TRUE;
           END_CASE;
       END_IF;
   END_IF;
END_FUNCTION

FUNCTION "Screens" : Void   // FC12, SCL
{ S7_Optimized_Access := 'TRUE' }
VERSION : 0.1
// stored: AutoNumber true, IsIECCheckEnabled false, SetENOAutomatically false, UDAEnableTagReadback false
BEGIN
   REGION MAIN
       IF "VTD_Automatic_Button" THEN
           "Control_DB".VTD_Control.Instruction.Mode_Change :=
           "Control_DB".ECnv_Control.Instruction.Mode_Change :=
           "Control_DB".LCnv_Control[1].Instruction.Mode_Change :=
           "Control_DB".LCnv_Control[2].Instruction.Mode_Change :=
           "Control_DB".LCnv_Control[3].Instruction.Mode_Change :=
           "Control_DB".LCnv_Control[1].Safety_Stop_Cnrl.Mode :=
           "Control_DB".LCnv_Control[2].Safety_Stop_Cnrl.Mode :=
           "Control_DB".LCnv_Control[3].Safety_Stop_Cnrl.Mode := 3;

           "Control_DB".VTD_Control.Instruction.Enable :=
           "Control_DB".ECnv_Control.Instruction.Enable :=
           "Control_DB".LCnv_Control[1].Instruction.Enable :=
           "Control_DB".LCnv_Control[2].Instruction.Enable :=
           "Control_DB".LCnv_Control[3].Instruction.Enable := TRUE;
       END_IF;

       IF "Carrousel_Automatic_Button" THEN
           "Control_DB".Inbound_Cnv.Instruction.Mode_Change :=
           "Control_DB".Outbound_Cnv.Instruction.Mode_Change :=
           "Control_DB".Pick_Station.Instruction.Mode_Change :=
           "Control_DB".PopUp_Cnv[1].Instruction.Mode_Change :=
           "Control_DB".PopUp_Cnv[2].Instruction.Mode_Change :=
           "Control_DB".PopUp_Cnv[3].Instruction.Mode_Change :=
           "Control_DB".PopUp_Cnv[4].Instruction.Mode_Change := 3;

           "Control_DB".Inbound_Cnv.Instruction.Enable :=
           "Control_DB".Outbound_Cnv.Instruction.Enable :=
           "Control_DB".Pick_Station.Instruction.Enable :=
           "Control_DB".PopUp_Cnv[1].Instruction.Enable :=
           "Control_DB".PopUp_Cnv[2].Instruction.Enable :=
           "Control_DB".PopUp_Cnv[3].Instruction.Enable :=
           "Control_DB".PopUp_Cnv[4].Instruction.Enable := TRUE;
       END_IF;

       "VTD_Buffers_In_Automatic" := "Control_DB".VTD_Control.Mode = 3 AND
       "Control_DB".ECnv_Control.Mode = 3 AND
       "Control_DB".LCnv_Control[1].Mode = 3 AND
       "Control_DB".LCnv_Control[2].Mode = 3 AND
       "Control_DB".LCnv_Control[3].Mode = 3 AND
       "Control_DB".LCnv_Control[1].Safety_Stop_Cnrl.Mode = 3 AND
       "Control_DB".LCnv_Control[2].Safety_Stop_Cnrl.Mode = 3 AND
       "Control_DB".LCnv_Control[3].Safety_Stop_Cnrl.Mode = 3;

       "Carrousel_In_Automatic" :=
       "Control_DB".Inbound_Cnv.Mode = 3 AND
       "Control_DB".Outbound_Cnv.Mode = 3 AND
       "Control_DB".Pick_Station.Mode = 3 AND
       "Control_DB".PopUp_Cnv[1].Mode = 3 AND
       "Control_DB".PopUp_Cnv[2].Mode = 3 AND
       "Control_DB".PopUp_Cnv[3].Mode = 3 AND
       "Control_DB".PopUp_Cnv[4].Mode = 3;

       IF "HMI_DB".ScreenNo = 0 THEN
           "Control_DB".VTD_Control.Instruction.Reset :=
           "Control_DB".ECnv_Control.Instruction.Reset :=
           "Control_DB".LCnv_Control[1].Instruction.Reset :=
           "Control_DB".LCnv_Control[2].Instruction.Reset :=
           "Control_DB".LCnv_Control[3].Instruction.Reset :=
           "Control_DB".Inbound_Cnv.Instruction.Reset :=
           "Control_DB".Outbound_Cnv.Instruction.Reset :=
           "Control_DB".Pick_Station.Instruction.Reset :=
           "Control_DB".PopUp_Cnv[1].Instruction.Reset :=
           "Control_DB".PopUp_Cnv[2].Instruction.Reset :=
           "Control_DB".PopUp_Cnv[3].Instruction.Reset :=
           "Control_DB".PopUp_Cnv[4].Instruction.Reset := "Reset_All";
       END_IF;

       //empty background
       IF "System_DB_VTD".Error OR "System_DB_Carousel".Error OR "Error_Word_1".%X0 THEN
           "Screen_DB".EmptyTemplate_Background := 1;
       ELSE
           "Screen_DB".EmptyTemplate_Background := 0;
       END_IF;

       //main background
       IF "HMI_DB".ScreenNo = 1 AND "System_DB_VTD".Error THEN
           "Screen_DB".MainTemplate_Background := 1;
       ELSIF "HMI_DB".ScreenNo = 2 AND "System_DB_Carousel".Error THEN
           "Screen_DB".MainTemplate_Background := 1;
       ELSIF "HMI_DB".ScreenNo <> 1 AND "HMI_DB".ScreenNo <> 2 AND ("System_DB_VTD".Error OR "System_DB_Carousel".Error OR "Error_Word_1".%X0) THEN
           "Screen_DB".MainTemplate_Background := 1;
       ELSE
           "Screen_DB".MainTemplate_Background := 0;
       END_IF;
   END_REGION 

   REGION SHUTTLES
       CASE "Screen_DB".Shuttle_Select OF
           1:
               "Screen_DB".Shuttle := "Shuttle_MQTT_DB".Shuttle_MQTT[1].Message.Shuttle_Status;
           2:
               "Screen_DB".Shuttle := "Shuttle_MQTT_DB".Shuttle_MQTT[2].Message.Shuttle_Status;
           3:
               "Screen_DB".Shuttle := "Shuttle_MQTT_DB".Shuttle_MQTT[3].Message.Shuttle_Status;
       END_CASE;
   END_REGION
END_FUNCTION

FUNCTION "GeneralErros_HMII" : Void   // FC13, SCL
{ S7_Optimized_Access := 'TRUE' }
VERSION : 0.1
// stored: AutoNumber true, IsIECCheckEnabled false, SetENOAutomatically false, UDAEnableTagReadback false
BEGIN
   "HMI_DB".GeneralErrors.%X0 := "Control_DB".LCnv_Control[1].Safety_Stop_Cnrl.Error;
   "HMI_DB".GeneralErrors.%X1 := "Control_DB".LCnv_Control[1].Safety_Stop_Cnrl.Error;
   "HMI_DB".GeneralErrors.%X2 := "Control_DB".LCnv_Control[2].Safety_Stop_Cnrl.Error;
   "HMI_DB".GeneralErrors.%X3 := "Control_DB".LCnv_Control[2].Safety_Stop_Cnrl.Error;
   "HMI_DB".GeneralErrors.%X4 := "Control_DB".LCnv_Control[3].Safety_Stop_Cnrl.Error;
   "HMI_DB".GeneralErrors.%X5 := "Control_DB".LCnv_Control[3].Safety_Stop_Cnrl.Error;

   "Error" := "System_DB_VTD".Error OR "System_DB_Carousel".Error;
END_FUNCTION

FUNCTION "FC_Orders" : Void   // FC96, SCL
{ S7_Optimized_Access := 'TRUE' }
VERSION : 0.1
// stored: AutoNumber true, IsIECCheckEnabled false, SetENOAutomatically false, UDAEnableTagReadback false
   VAR_TEMP
      i : Int;
      j : Int;
      EmptyOrder : "OrderTable_UDT";
   END_VAR
BEGIN
   //Main Screen
   //IF "HMI_DB".ScreenNo = 1 THEN
       FOR #i := 1 TO 5 DO
           "HMI_OrderTable".Index_1[#i] := #i;
           "HMI_OrderTable".OrderTable_1[#i] := "System_DB_Carousel".OrderTable[#i];
           "HMI_OrderTable".Index_2[#i] := #i;
           "HMI_OrderTable".OrderTable_2[#i] := "System_DB_VTD".OrderTable[#i];

           //Color State
           IF "HMI_OrderTable".OrderTable_1[#i].Status = 'Queued' THEN
               "HMI_OrderTable".State_1[#i] := 1;
           ELSIF "HMI_OrderTable".OrderTable_1[#i].Status = 'Running' THEN
               "HMI_OrderTable".State_1[#i] := 2;
           ELSIF "HMI_OrderTable".OrderTable_1[#i].Status = 'Completed' THEN
               "HMI_OrderTable".State_1[#i] := 3;
           ELSIF "HMI_OrderTable".OrderTable_1[#i].Status = 'Error' THEN
               "HMI_OrderTable".State_1[#i] := 4;
           ELSIF "HMI_OrderTable".OrderTable_1[#i].Status = 'Paused' THEN
               "HMI_OrderTable".State_1[#i] := 5;
           ELSIF "HMI_OrderTable".OrderTable_1[#i].Status = 'Canceled' THEN
               "HMI_OrderTable".State_1[#i] := 6;
           ELSIF "HMI_OrderTable".OrderTable_1[#i].Status = 'Error\Cancel' THEN
               "HMI_OrderTable".State_1[#i] := 7;
           ELSE
               "HMI_OrderTable".State_1[#i] := 0;
           END_IF;

           IF "HMI_OrderTable".OrderTable_2[#i].Status = 'Queued' THEN
               "HMI_OrderTable".State_2[#i] := 1;
           ELSIF "HMI_OrderTable".OrderTable_2[#i].Status = 'Running' THEN
               "HMI_OrderTable".State_2[#i] := 2;
           ELSIF "HMI_OrderTable".OrderTable_2[#i].Status = 'Completed' THEN
               "HMI_OrderTable".State_2[#i] := 3;
           ELSIF "HMI_OrderTable".OrderTable_2[#i].Status = 'Error' THEN
               "HMI_OrderTable".State_2[#i] := 4;
           ELSIF "HMI_OrderTable".OrderTable_2[#i].Status = 'Paused' THEN
               "HMI_OrderTable".State_2[#i] := 5;
           ELSIF "HMI_OrderTable".OrderTable_2[#i].Status = 'Canceled' THEN
               "HMI_OrderTable".State_2[#i] := 6;
           ELSIF "HMI_OrderTable".OrderTable_2[#i].Status = 'Error\Cancel' THEN
               "HMI_OrderTable".State_2[#i] := 7;
           ELSE
               "HMI_OrderTable".State_2[#i] := 0;
           END_IF;

       END_FOR;
   //END_IF;

   IF "HMI_OrderTable".StartRow < 0 THEN
       "HMI_OrderTable".StartRow := 0;
   END_IF;
   IF "HMI_OrderTable".StartRow > 90 THEN
       "HMI_OrderTable".StartRow := 90;
   END_IF;

   //System #1 - Carousel Order Table
   //IF "HMI_DB".ScreenNo = 407 AND "HMI_Systems".SystemNo = 1 THEN
           //Place New Order manually
       IF "HMI_OrderTable".PlaceOrder_PB  AND "HMI_OrderTable".PlacingNewOrder THEN
           "HMI_OrderTable".PlaceOrder_PB := FALSE;
           CASE "HMI_OrderTable".Device OF
               1:
                   "HMI_OrderTable".OrderTable_1[0].Device := 'Roller to Roller'; //6
               3:
                   "HMI_OrderTable".OrderTable_1[0].Device := 'Chain to Chain'; //7
               5:
                   "HMI_OrderTable".OrderTable_1[0].Device := 'Pop4 to Pick';//8
               6:
                   "HMI_OrderTable".OrderTable_1[0].Device := 'Pick to Pop1';//9
               7:
                   "HMI_OrderTable".OrderTable_1[0].Device := 'Weigh Station';//10
               9:
                   "HMI_OrderTable".OrderTable_1[0].Device := 'Profile Station';//14
               // 10:
               //     "HMI_OrderTable".OrderTable_1[0].Device := 'LB Exit 1';
               // 11:
               //     "HMI_OrderTable".OrderTable_1[0].Device := 'CM 1';

           END_CASE;
           IF "HMI_OrderTable".Device > 9 THEN
               "HMI_OrderTable".OrderTable_1[0].OPC_Control.Destination_Location := 0;
           END_IF;
          // "System_DB_Carousel".OrderSent := "HMI_OrderTable".Device > 0;
           "System_DB_Carousel".StepTable[1] := "HMI_OrderTable".OrderTable_1[0];
           "System_DB_Carousel".StepTable[1].OrderNo := -1;
           "System_DB_Carousel".StepTable[1].StepNo := -1;
           "System_DB_Carousel".StepTable[1].PlaceTime := "Time".CurrentLocalTime;
           "System_DB_Carousel".StepTable[1].Status := 'Queued';
       END_IF;

       //Pause Order Push Button
       IF "HMI_OrderTable".PauseOrders_PB THEN
           "HMI_OrderTable".PauseOrders_PB := FALSE;
           "System_DB_Carousel".PauseOrders := TRUE;
       END_IF;
       //Resume Order Push Button
       IF "HMI_OrderTable".ResumeOrder_PB THEN
           "HMI_OrderTable".ResumeOrder_PB := FALSE;
           "System_DB_Carousel".ResumeOrders := TRUE;
       END_IF;
       //Cancel Order Push Button
       IF "HMI_OrderTable".CancelOrder_PB THEN
           "HMI_OrderTable".CancelOrder_PB := FALSE;
           "System_DB_Carousel".CancelOrders := TRUE;
       END_IF;
       //Cancel This Order Push Button
       IF "HMI_OrderTable".CancelThisOrder_PB THEN
           "HMI_OrderTable".CancelThisOrder_PB := FALSE;
           IF "HMI_OrderTable".OrderTable_1["HMI_OrderTable".PopUp_Index].Status = 'Error' THEN
               "System_DB_Carousel".OrderTable["HMI_OrderTable".PopUp_Index + "HMI_OrderTable".StartRow].Status := 'Error\Cancel';
               IF "System_DB_Carousel".CurrentOrder = "HMI_OrderTable".PopUp_Index THEN
                   "System_DB_Carousel".CurrentOrder -= 1;
               END_IF;
               IF "System_DB_Carousel".OrderTable["HMI_OrderTable".PopUp_Index + "HMI_OrderTable".StartRow].Device = 'Roller to Roller' THEN
                   "System_Unit_1".Roller_To_Roller_CurrentOrder := 0;
               ELSIF "System_DB_Carousel".OrderTable["HMI_OrderTable".PopUp_Index + "HMI_OrderTable".StartRow].Device = 'Chain to Chain' THEN
                   "System_Unit_1".Chain_To_Chain_CurrentOrder := 0;
               ELSIF "System_DB_Carousel".OrderTable["HMI_OrderTable".PopUp_Index + "HMI_OrderTable".StartRow].Device = 'Pop4 to Pick' THEN
                   "System_Unit_1".Pop4_To_PickSt_CurrentOrder := 0;
               ELSIF "System_DB_Carousel".OrderTable["HMI_OrderTable".PopUp_Index + "HMI_OrderTable".StartRow].Device = 'Pick to Pop1' THEN
                   "System_Unit_1".PickSt_To_Pop1_CurrentOrder := 0;
               ELSIF "System_DB_Carousel".OrderTable["HMI_OrderTable".PopUp_Index + "HMI_OrderTable".StartRow].Device = 'Weigh Station' THEN
                   "System_Unit_1".WeighingStation_CurrentOrder := 0;
               ELSIF "System_DB_Carousel".OrderTable["HMI_OrderTable".PopUp_Index + "HMI_OrderTable".StartRow].Device = 'Profile Station' THEN
                   "System_Unit_1".ProfileStation_CurrentOrder := 0;

               END_IF;
           END_IF;

       END_IF;

       //Copy data
       FOR #i := 1 TO 9 DO
           #j := "HMI_OrderTable".StartRow + #i;
           "HMI_OrderTable".Index_1[#i] := #j;
           "HMI_OrderTable".OrderTable_1[#i] := "System_DB_Carousel".OrderTable[#j];
                   //Color State
           IF "HMI_OrderTable".OrderTable_1[#i].Status = 'Queued' THEN
               "HMI_OrderTable".State_1[#i] := 1;
           ELSIF "HMI_OrderTable".OrderTable_1[#i].Status = 'Running' THEN
               "HMI_OrderTable".State_1[#i] := 2;
           ELSIF "HMI_OrderTable".OrderTable_1[#i].Status = 'Completed' THEN
               "HMI_OrderTable".State_1[#i] := 3;
           ELSIF "HMI_OrderTable".OrderTable_1[#i].Status = 'Error' THEN
               "HMI_OrderTable".State_1[#i] := 4;
           ELSIF "HMI_OrderTable".OrderTable_1[#i].Status = 'Paused' THEN
               "HMI_OrderTable".State_1[#i] := 5;
           ELSIF "HMI_OrderTable".OrderTable_1[#i].Status = 'Canceled' THEN
               "HMI_OrderTable".State_1[#i] := 6;
           ELSIF "HMI_OrderTable".OrderTable_1[#i].Status = 'Error\Cancel' THEN
               "HMI_OrderTable".State_1[#i] := 7;
           ELSE
               "HMI_OrderTable".State_1[#i] := 0;
           END_IF;
       END_FOR;
   //END_IF;


   //System #2 - VTD Order Table
   //IF "HMI_DB".ScreenNo = 407 AND  "HMI_Systems".SystemNo= 2 THEN

       //Place Order manually
       IF "HMI_OrderTable".PlaceOrder_PB AND "HMI_OrderTable".PlacingNewOrder THEN
           "HMI_OrderTable".PlaceOrder_PB := FALSE;
           CASE "HMI_OrderTable".Device OF

               1:
                   "HMI_OrderTable".OrderTable_2[0].Device := 'VTD';
               2:
                   "HMI_OrderTable".OrderTable_2[0].Device := 'Pallet In Out';
               3:
                   "HMI_OrderTable".OrderTable_2[0].Device := 'Shuttle In Out';
               // 4:
               //     "HMI_OrderTable".OrderTable_1[0].Device := 'Shuttle 2';
               // 5:
               //     "HMI_OrderTable".OrderTable_1[0].Device := 'TurnTable';
               // 6:
               //     "HMI_OrderTable".OrderTable_1[0].Device := 'LS VRC 2';
               // 7:
               //     "HMI_OrderTable".OrderTable_1[0].Device := 'HS VRC 1';
               // 8:
               //     "HMI_OrderTable".OrderTable_1[0].Device := 'HS VRC 2';
               // 9:
               //     "HMI_OrderTable".OrderTable_1[0].Device := 'LB Entry 2';
               // 10:
               //     "HMI_OrderTable".OrderTable_1[0].Device := 'LB Exit 2';
               // 11:
               //     "HMI_OrderTable".OrderTable_1[0].Device := 'CM 2';


           END_CASE;
           IF "HMI_OrderTable".Device > 9 THEN
               "HMI_OrderTable".OrderTable_2[0].OPC_Control.Destination_Location := 0;
           END_IF;
          // "System_DB_VTD".OrderSent := "HMI_OrderTable".Device > 0;
           "System_DB_VTD".StepTable[1] := "HMI_OrderTable".OrderTable_2[0];
           "System_DB_VTD".StepTable[1].OrderNo := -1;
           "System_DB_VTD".StepTable[1].StepNo := -1;
           "System_DB_VTD".StepTable[1].PlaceTime := "Time".CurrentLocalTime;
           "System_DB_VTD".StepTable[1].Status := 'Queued';
       END_IF;

       //Pause Order Push Button
       IF "HMI_OrderTable".PauseOrders_PB THEN
           "HMI_OrderTable".PauseOrders_PB := FALSE;
           "System_DB_VTD".PauseOrders := TRUE;
       END_IF;
       //Resume Order Push Button
       IF "HMI_OrderTable".ResumeOrder_PB THEN
           "HMI_OrderTable".ResumeOrder_PB := FALSE;
           "System_DB_VTD".ResumeOrders := TRUE;
       END_IF;
       //Cancel Order Push Button
       IF "HMI_OrderTable".CancelOrder_PB THEN
           "HMI_OrderTable".CancelOrder_PB := FALSE;
           "System_DB_VTD".CancelOrders := TRUE;
       END_IF;

       //Cancel This Order Push Button
       IF "HMI_OrderTable".CancelThisOrder_PB THEN
           "HMI_OrderTable".CancelThisOrder_PB := FALSE;
           IF "HMI_OrderTable".OrderTable_2["HMI_OrderTable".PopUp_Index].Status = 'Error' THEN
               "System_DB_VTD".OrderTable["HMI_OrderTable".PopUp_Index].Status := 'Error\Cancel';
               IF "System_DB_VTD".CurrentOrder = "HMI_OrderTable".PopUp_Index THEN
                   "System_DB_VTD".CurrentOrder -= 1;
               END_IF;


               IF "System_DB_VTD".OrderTable["HMI_OrderTable".PopUp_Index + "HMI_OrderTable".StartRow].Device = 'VTD' THEN
                   "System_Unit_2".VTD_CurrentOrder := 0;
               ELSIF "System_DB_VTD".OrderTable["HMI_OrderTable".PopUp_Index + "HMI_OrderTable".StartRow].Device = 'Pallet In Out' THEN
                   "System_Unit_2".Pallet_InOut_CurrentOrder := 0;
               ELSIF "System_DB_VTD".OrderTable["HMI_OrderTable".PopUp_Index + "HMI_OrderTable".StartRow].Device = 'Shuttle In Out' THEN
                   "System_Unit_2".Shuttle_InOut_CurrentOrder := 0;
                   // ELSIF "System_DB_VTD".OrderTable["HMI_OrderTable".PopUp_Index + "HMI_OrderTable".StartRow].Device = 'Shuttle 2' THEN
                   //     "System_Unit_2".Shuttle_2_CurrentOrder := 0;
                   // ELSIF "System_DB_VTD".OrderTable["HMI_OrderTable".PopUp_Index + "HMI_OrderTable".StartRow].Device = 'TurnTable' THEN
                   //     "System_Unit_2".TurnTable_CurrentOrder := 0;
                   // ELSIF "System_DB_VTD".OrderTable["HMI_OrderTable".PopUp_Index + "HMI_OrderTable".StartRow].Device = 'HS VRC 1' THEN
                   //     "System_Unit_2".HS_VRC_1_CurrentOrder := 0;
                   // ELSIF "System_DB_VTD".OrderTable["HMI_OrderTable".PopUp_Index + "HMI_OrderTable".StartRow].Device = 'HS VRC 2' THEN
                   //     "System_Unit_2".HS_VRC_2_CurrentOrder := 0;
                   // ELSIF "System_DB_VTD".OrderTable["HMI_OrderTable".PopUp_Index + "HMI_OrderTable".StartRow].Device = 'LB Entry 2' THEN
                   //     "System_Unit_2".LoadingBayEntry_2_CurrentOrder := 0;
                   // ELSIF "System_DB_VTD".OrderTable["HMI_OrderTable".PopUp_Index + "HMI_OrderTable".StartRow].Device = 'LB Exit 2' THEN
                   //     "System_Unit_2".LoadingBayExit_2_CurrentOrder := 0;
                   // ELSIF "System_DB_VTD".OrderTable["HMI_OrderTable".PopUp_Index + "HMI_OrderTable".StartRow].Device = 'LS VRC 2' THEN
                   //     "System_Unit_2".LS_VRC_2_CurrentOrder := 0;

               END_IF;

           END_IF;

       END_IF;

       //Copy data
       FOR #i := 1 TO 9 DO
           #j := "HMI_OrderTable".StartRow + #i;
           "HMI_OrderTable".Index_2[#i] := #j;
           "HMI_OrderTable".OrderTable_2[#i] := "System_DB_VTD".OrderTable[#j];
           //Color State
           IF "HMI_OrderTable".OrderTable_2[#i].Status = 'Queued' THEN
               "HMI_OrderTable".State_2[#i] := 1;
           ELSIF "HMI_OrderTable".OrderTable_2[#i].Status = 'Running' THEN
               "HMI_OrderTable".State_2[#i] := 2;
           ELSIF "HMI_OrderTable".OrderTable_2[#i].Status = 'Completed' THEN
               "HMI_OrderTable".State_2[#i] := 3;
           ELSIF "HMI_OrderTable".OrderTable_2[#i].Status = 'Error' THEN
               "HMI_OrderTable".State_2[#i] := 4;
           ELSIF "HMI_OrderTable".OrderTable_2[#i].Status = 'Paused' THEN
               "HMI_OrderTable".State_2[#i] := 5;
           ELSIF "HMI_OrderTable".OrderTable_2[#i].Status = 'Canceled' THEN
               "HMI_OrderTable".State_2[#i] := 6;
           ELSIF "HMI_OrderTable".OrderTable_2[#i].Status = 'Error\Cancel' THEN
               "HMI_OrderTable".State_2[#i] := 7;
           ELSE
               "HMI_OrderTable".State_2[#i] := 0;
           END_IF;
       END_FOR;
   //END_IF;



   IF NOT "HMI_OrderTable".PlacingNewOrder THEN
       "HMI_OrderTable".Device := 0;
   END_IF;

   //Error PopUp Window
   IF "HMI_OrderTable".PopUp_ErrorWindow_Active AND NOT "HMI_OrderTable".PlacingNewOrder THEN
       "HMI_OrderTable".OrderTable_2[0] := "HMI_OrderTable".OrderTable_2["HMI_OrderTable".PopUp_Index];
       IF "HMI_OrderTable".OrderTable_2[0].Status = 'Error' THEN
           "HMI_OrderTable".State_2[0] := 4;
       ELSIF "HMI_OrderTable".OrderTable_2[0].Status = 'Error\Cancel' THEN
           "HMI_OrderTable".State_2[0] := 7;
       ELSE
           "HMI_OrderTable".State_2[0] := 0;
       END_IF;
   ELSIF NOT "HMI_OrderTable".PopUp_ErrorWindow_Active AND NOT "HMI_OrderTable".PlacingNewOrder THEN
       "HMI_OrderTable".OrderTable_2[0] := #EmptyOrder;
   END_IF;
END_FUNCTION

FUNCTION "Errors" : Void   // FC26, SCL
{ S7_Optimized_Access := 'TRUE' }
VERSION : 0.1
// stored: AutoNumber true, IsIECCheckEnabled false, SetENOAutomatically false, UDAEnableTagReadback false
   VAR_TEMP
      ReturnValue : Word;
      Devices : Array[0..1023] of Bool;
   END_VAR
BEGIN
   REGION Profinet Device Errors
       #ReturnValue := DeviceStates(LADDR := "Local~PROFINET_IO-System",
                                    MODE := 2, // Mode 5 = a problem has occurred
                                    STATE := #Devices);
       IF #ReturnValue = 0 THEN
           IF #Devices[0] THEN // Main PLC Error
               "Errors_Profinet_1".%X0 := TRUE;
           END_IF;

           IF #Devices[1] THEN // Switch 1
               "Errors_Profinet_1".%X1 := TRUE;
           END_IF;

           IF #Devices[2] THEN // Switch 2
               "Errors_Profinet_1".%X2 := TRUE;
           END_IF;

           IF #Devices[3] THEN // Remote IO
               "Errors_Profinet_1".%X3 := TRUE;
           END_IF;

           IF #Devices[4] THEN // VTD
               "Errors_Profinet_1".%X4 := TRUE;
           END_IF;

           IF #Devices[5] THEN // Lift PopUp1
               "Errors_Profinet_1".%X5 := TRUE;
           END_IF;

           IF #Devices[6] THEN // Lift PopUp4
               "Errors_Profinet_1".%X6 := TRUE;
           END_IF;

           IF #Devices[7] THEN // Lift PopUp2
               "Errors_Profinet_1".%X7 := TRUE;
           END_IF;

           IF #Devices[8] THEN // Roller Outbound
               "Errors_Profinet_1".%X8 := TRUE;
           END_IF;

           IF #Devices[9] THEN // Roller Inbound
               "Errors_Profinet_1".%X9 := TRUE;
           END_IF;

           IF #Devices[10] THEN // Roller PopUp1
               "Errors_Profinet_1".%X10 := TRUE;
           END_IF;

           IF #Devices[11] THEN // Roller PopUp2
               "Errors_Profinet_1".%X11 := TRUE;
           END_IF;

           IF #Devices[12] THEN // Roller PopUp3
               "Errors_Profinet_1".%X12 := TRUE;
           END_IF;

           IF #Devices[13] THEN // Chain 1
               "Errors_Profinet_1".%X13 := TRUE;
           END_IF;

           IF #Devices[14] THEN // Chain 2
               "Errors_Profinet_1".%X14 := TRUE;
           END_IF;

           IF #Devices[15] THEN // Chain 3
               "Errors_Profinet_1".%X15 := TRUE;
           END_IF;

           IF #Devices[16] THEN // Buffer Level 1
               "Errors_Profinet_2".%X0 := TRUE;
           END_IF;

           IF #Devices[17] THEN // Buffer Level 2
               "Errors_Profinet_2".%X1 := TRUE;
           END_IF;

           IF #Devices[18] THEN // Buffer Level 3
               "Errors_Profinet_2".%X2 := TRUE;
           END_IF;

           IF #Devices[19] THEN // Roller PopUp4
               "Errors_Profinet_2".%X3 := TRUE;
           END_IF;

           IF #Devices[20] THEN // VTD Conveyor
               "Errors_Profinet_2".%X4 := TRUE;
           END_IF;

           IF #Devices[21] THEN // IND360
               "Errors_Profinet_2".%X5 := TRUE;
           END_IF;

           IF #Devices[22] THEN // Lift PopUp3
               "Errors_Profinet_2".%X6 := TRUE;
           END_IF;

           IF #Devices[23] THEN // Turck
               "Errors_Profinet_2".%X7 := TRUE;
           END_IF;

           IF #Devices[24] THEN // INTERFACE ET200AL
               "Errors_Profinet_2".%X8 := TRUE;
           END_IF;

           IF #Devices[25] THEN // WLAN 1
               "Errors_Profinet_2".%X9 := TRUE;
           END_IF;

           IF #Devices[26] THEN // WLAN 2
               "Errors_Profinet_2".%X10 := TRUE;
           END_IF;

           IF #Devices[27] THEN // WLAN 3
               "Errors_Profinet_2".%X11 := TRUE;
           END_IF;

           IF #Devices[28] THEN // WLAN 4
               "Errors_Profinet_2".%X12 := TRUE;
           END_IF;

           IF #Devices[29] THEN // Linear Encoder
               "Errors_Profinet_2".%X13 := TRUE;
           END_IF;

           IF #Devices[30] THEN // Absolute Encoder
               "Errors_Profinet_2".%X14 := TRUE;
           END_IF;

           IF #Devices[31] THEN // Sick Barcode
               "Errors_Profinet_2".%X15 := TRUE;
           END_IF;

           IF #Devices[32] THEN // Inbound Leuze Barcode
               "Errors_Profinet_3".%X0 := TRUE;
           END_IF;

           IF #Devices[33] THEN // Outbound Leuze Barcode
               "Errors_Profinet_3".%X1 := TRUE;
           END_IF;

           IF #Devices[34] THEN // HMI
               "Errors_Profinet_3".%X2 := TRUE;
           END_IF;

           IF #Devices[35] THEN // Light Guard
               "Errors_Profinet_3".%X3 := TRUE;
           END_IF;
       END_IF;
   END_REGION

   REGION LMs
       IF NOT "Auxiliar Circuit Breaker Feedback LM2" THEN
           "Erros_LMs_1".%X0 := TRUE;
       END_IF;

       IF NOT "Auxiliar Circuit Breaker Feedback LM3" THEN
           "Erros_LMs_1".%X1 := TRUE;
       END_IF;

       IF NOT "Auxiliar Circuit Breaker Feedback LM4" THEN
           "Erros_LMs_1".%X2 := TRUE;
       END_IF;

       IF NOT "Auxiliar Circuit Breaker Feedback LM5" THEN
           "Erros_LMs_1".%X3 := TRUE;
       END_IF;

       IF NOT "Auxiliar Circuit Breaker Feedback LM6" THEN
           "Erros_LMs_1".%X4 := TRUE;
       END_IF;

       IF NOT "Auxiliar Circuit Breaker Feedback LM7" THEN
           "Erros_LMs_1".%X5 := TRUE;
       END_IF;

       IF NOT "Auxiliar Circuit Breaker Feedback LM8" THEN
           "Erros_LMs_1".%X6 := TRUE;
       END_IF;

       IF NOT "Auxiliar Circuit Breaker Feedback LM9" THEN
           "Erros_LMs_1".%X7 := TRUE;
       END_IF;

       IF NOT "Auxiliar Circuit Breaker Feedback LM10" THEN
           "Erros_LMs_1".%X8 := TRUE;
       END_IF;

       IF NOT "Auxiliar Circuit Breaker Feedback LM11" THEN
           "Erros_LMs_1".%X9 := TRUE;
       END_IF;

       IF NOT "Auxiliar Circuit Breaker Feedback LM12" THEN
           "Erros_LMs_1".%X10 := TRUE;
       END_IF;

       IF NOT "Auxiliar Circuit Breaker Feedback LM13" THEN
           "Erros_LMs_1".%X11 := TRUE;
       END_IF;

       IF NOT "Auxiliar Circuit Breaker Feedback LM14" THEN
           "Erros_LMs_1".%X12 := TRUE;
       END_IF;

       IF NOT "Auxiliar Circuit Breaker Feedback LM15" THEN
           "Erros_LMs_1".%X13 := TRUE;
       END_IF;

       IF NOT "Auxiliar Circuit Breaker Feedback LM16" THEN
           "Erros_LMs_1".%X14 := TRUE;
       END_IF;

       IF NOT "Auxiliar Circuit Breaker Feedback LM100" THEN
           "Erros_LMs_1".%X15 := TRUE;
       END_IF;

       IF NOT "Auxiliar Circuit Breaker Feedback LM101" THEN
           "Erros_LMs_2".%X0 := TRUE;
       END_IF;

       IF NOT "Auxiliar Circuit Breaker Feedback LM102" THEN
           "Erros_LMs_2".%X1 := TRUE;
       END_IF;

       IF NOT "Auxiliar Circuit Breaker Feedback LM103" THEN
           "Erros_LMs_2".%X2 := TRUE;
       END_IF;

       IF NOT "Auxiliar Circuit Breaker Feedback LM104" THEN
           "Erros_LMs_2".%X3 := TRUE;
       END_IF;

       IF NOT "Auxiliar Circuit Breaker Feedback LM105" THEN
           "Erros_LMs_2".%X4 := TRUE;
       END_IF;

       IF NOT "Auxiliar Circuit Breaker Feedback LM106" THEN
           "Erros_LMs_2".%X5 := TRUE;
       END_IF;

       IF NOT "Auxiliar Circuit Breaker Feedback LM107" THEN
           "Erros_LMs_2".%X6 := TRUE;
       END_IF;

   END_REGION

   REGION WEIGHT STATION
       REGION Smart5 Red Level 5 

           // Calibration error 
           "Errors_IND360_Smart5_Red_Level_5".%X0 := "SB Status Group 1".%X0;
           // 1 = Weight data can no longer be trusted
           // due TO loss OF calibration data OR an
           // algorithm running in the product TO detect
           // weighing irregularities.

           // Out of A/D range over/under
           "Errors_IND360_Smart5_Red_Level_5".%X1 := "SB Status Group 1".%X1;
           // 1 = Weight data can no longer be trusted
           // due TO loss OF data OR mechanical damage
           // OF the weigh module.

           // Checksum failure 
           "Errors_IND360_Smart5_Red_Level_5".%X2 := "SB Status Group 1".%X2;
           // 1 = A checksum analysis OF memory does
           // NOT yield the expected result.

           // Weight blocked
           "Errors_IND360_Smart5_Red_Level_5".%X3 := "SB Status Group 1".%X3;
           // [NOT supported BY IND360 devices.]

           // Single sensor communication failure (LC missing)
           "Errors_IND360_Smart5_Red_Level_5".%X4 := "SB Status Group 1".%X4;
           // 1 = One OR more OF the connected sensors
           // are NOT working properly.

           //Customer defined overload
           "Errors_IND360_Smart5_Red_Level_5".%X5 := "SB Status Group 1".%X5;
           // 1 = Weight is equal TO OR greater than the
           // maximum load allowed. Although overload
           // is a conditional limit, it can lead TO bigger
           // #Errors such as mechanical breakage OR
           // personal injury.

           // Customer defined underload
           "Errors_IND360_Smart5_Red_Level_5".%X6 := "SB Status Group 1".%X6;
           // 1 = Weight is equal OR less than the
           // minimum load allowed.

           // Network failure (all cells)
           "Errors_IND360_Smart5_Red_Level_5".%X7 := "SB Status Group 1".%X7;
           // Applicable only on multi-cell networks.
           // 1 = Failure OF the entire Network. No cells
           // are responding.

           // Zero out OF range
           "Errors_IND360_Smart5_Red_Level_5".%X8 := "SB Status Group 1".%X8;
           // 1 = A control system attempted A Zero
           // command but the device did NOT accept the
           // command because the weight is outside the
           // specified limits OR the weights AND measure
           // limits.

           // Symmetry #Errors
           "Errors_IND360_Smart5_Red_Level_5".%X9 := "SB Status Group 1".%X9;
           // Applicable only FOR products with TraxDSP
           // function which detects significant errors
           // between load cells AND their peers.
           // 1 = A symmetry error has been detected.

           // Temperature #Errors (LC temperature out OF normal temperature)
           "Errors_IND360_Smart5_Red_Level_5".%X10 := "SB Status Group 1".%X10;
           // 1 = Sensor is outside OF the allowed
           // Temperature range. The weight value can be
           // affected, OR the components can prematurely
           // fail.

           // Weights AND measures failure
           "Errors_IND360_Smart5_Red_Level_5".%X11 := "SB Status Group 1".%X11;
           // 1 = The product is no longer in compliance
           // with Weights AND measure regulations.

           // Foreign device detected
           "Errors_IND360_Smart5_Red_Level_5".%X12 := "SB Status Group 1".%X12;
           // 1 = A Foreign device is attached TO the
           // system OR any similar algorithm limits.

           // Test mode
           "Errors_IND360_Smart5_Red_Level_5".%X13 := "SB Status Group 1".%X13;
           // 1 = Device is in a mode in which live data
           // is being replaced with special Test data.

           // Analog LC Error
           "Errors_IND360_Smart5_Red_Level_5".%X14 := "SB Status Group 1".%X14;
           // 1 = Analog Sensor Error detected BY
           // measuring system total resistance
       END_REGION
   END_REGION

   REGION Leuze Barcode
       //INBOUND LECTOR
       IF "In Lector_Staus" = 128 THEN
           "Error_Devices".%X0 := TRUE;
       ELSIF "In Lector_Staus" = 129 THEN
           "Error_Devices".%X1 := TRUE;
       END_IF;

       //OUTBOUND LECTOR
       IF "Out Lector_Staus" = 128 THEN
           "Error_Devices".%X2 := TRUE;
       ELSIF "Out Lector_Staus" = 129 THEN
           "Error_Devices".%X3 := TRUE;
       END_IF;
   END_REGION

   REGION Sick Barcode
       IF "SICK_Lector".Errorcode = 16#0000_0001 THEN //Timeout (SICK_CCOM_PNDP) 
           "Sick Lector_Error code 1".%X0 := TRUE;
       ELSIF "SICK_Lector".Errorcode = 16#0000_0002 THEN //Invalid module length (input)
           "Sick Lector_Error code 1".%X1 := TRUE;
       ELSIF "SICK_Lector".Errorcode = 16#0000_0003 THEN //Invalid module length (output)
           "Sick Lector_Error code 1".%X2 := TRUE;
       ELSIF "SICK_Lector".Errorcode = 16#0000_0004 THEN //DPWR_DAT error 
           "Sick Lector_Error code 1".%X3 := TRUE;
       ELSIF "SICK_Lector".Errorcode = 16#0000_0005 THEN //DPRD_DAT error 
           "Sick Lector_Error code 1".%X4 := TRUE;
       ELSIF "SICK_Lector".Errorcode > 16#0000_0006 AND "SICK_Lector".Errorcode < 16#0000_0009 THEN //Communication error 
           "Sick Lector_Error code 1".%X5 := TRUE;
       ELSIF "SICK_Lector".Errorcode = 16#0000_0010 THEN //Timeout (SICK_CCOM_PNDP)
           "Sick Lector_Error code 1".%X6 := TRUE;
       ELSIF "SICK_Lector".Errorcode = 16#0000_0011 THEN //Device error 
           "Sick Lector_Error code 1".%X7 := TRUE;
       ELSIF "SICK_Lector".Errorcode = 16#0000_0012 THEN //SICK_GetValue error 
           "Sick Lector_Error code 1".%X8 := TRUE;
       ELSIF "SICK_Lector".Errorcode = 16#0000_0013 THEN //SICK_SetValue error
           "Sick Lector_Error code 1".%X9 := TRUE;
       ELSIF "SICK_Lector".Errorcode = 16#0000_0014 THEN //#CANId > 63 
           "Sick Lector_Error code 1".%X10 := TRUE;
       ELSIF "SICK_Lector".Errorcode = 16#0000_0015 THEN //No module function selected, OR more than one module function selected
           "Sick Lector_Error code 1".%X11 := TRUE;
       ELSIF "SICK_Lector".Errorcode = 16#0000_0016 THEN //Invalid command response received
           "Sick Lector_Error code 1".%X12 := TRUE;
       ELSIF "SICK_Lector".Errorcode = 16#0000_0017 THEN //Change not possible in "RUN mode".
           "Sick Lector_Error code 1".%X13 := TRUE;
       ELSIF "SICK_Lector".Errorcode = 16#0000_0020 THEN //FreeCommand.sCommand > arrCommand (500 bytes)
           "Sick Lector_Error code 1".%X14 := TRUE;
       ELSIF "SICK_Lector".Errorcode = 16#0000_0021 THEN //Response to free command > result string(FreeCommand.sResult[100 characters])
           "Sick Lector_Error code 1".%X15 := TRUE;
       ELSIF "SICK_Lector".Errorcode = 16#0000_0022 THEN //String length Match - code.sName =0
           "Sick Lector_Error code 2".%X0 := TRUE;
       END_IF;
       END_REGION

   REGION Linear Encoder
       IF "LE_Status".%X0 THEN //Error present
           IF "LE_X_Unsafe_Position" = 1 THEN //Reader tilted 180°
               "Linear Encoder_Device Errors".%X0 := TRUE;
           ELSIF "LE_X_Unsafe_Position" = 2 THEN // No clear position can be determined (difference between codes is too great, code distance incorrect, etc.)
               "Linear Encoder_Device Errors".%X1 := TRUE;
           ELSIF "LE_X_Unsafe_Position" = 1000 THEN //Internal error
               "Linear Encoder_Device Errors".%X2 := TRUE;
           END_IF;
       ELSIF "LE_Status".%X1 THEN // No position information/OUT
           "Linear Encoder_Device Errors".%X3 := TRUE;
       ELSE//NO ERROR
           "Linear Encoder_Device Errors" := 0;
       END_IF;

       //WARNINGS
       IF "LE_Status".%X2 THEN // Warnign present
           "Linear Encoder_Warnings".%X0 := "LE_Warnings".%X0; //Code with non-PXV content found
           "Linear Encoder_Warnings".%X1 := "LE_Warnings".%X1; //Reader too close to code tape
           "Linear Encoder_Warnings".%X2 := "LE_Warnings".%X2; //Reader too far from code tape
           "Linear Encoder_Warnings".%X3 := "LE_Warnings".%X3; //Y position too large; the sensor is just before OUT
           "Linear Encoder_Warnings".%X4 := "LE_Warnings".%X4; //Y position too small; the sensor is just before OUT
           "Linear Encoder_Warnings".%X5 := "LE_Warnings".%X5; //The reader is rotated or tilted in relation to the code tape
           "Linear Encoder_Warnings".%X6 := "LE_Warnings".%X6; // Low level of code contrast
           "Linear Encoder_Warnings".%X7 := "LE_Warnings".%X7; //Repair tape detected
           "Linear Encoder_Warnings".%X8 := "LE_Warnings".%X8; //Temperature too high
           END_IF;
   END_REGION

   REGION RESET
       IF "Reset_All" THEN
           "Errors_Profinet_1" := 0;
           "Errors_Profinet_2" := 0;
           "Errors_Profinet_3" := 0;
           "Error_Devices" := 0;
           "Sick Lector_Error code 1" := 0;
           "Sick Lector_Error code 2" := 0;
           "Erros_LMs_1" := "Erros_LMs_2" := 0;
           "Linear Encoder_Device Errors" := 0;
       END_IF;
   END_REGION
END_FUNCTION

FUNCTION_BLOCK "InConveyor_FB"   // FB9, SCL
TITLE = Conveyor Instance FB
{ S7_Optimized_Access := 'TRUE' }
AUTHOR : Mertin Coetzee
VERSION : 0.1
// stored: AutoNumber true, IsIECCheckEnabled false, IsRetainMemResEnabled false, MemoryReserve 100, SetENOAutomatically false, UDAEnableTagReadback false
   VAR_INPUT
      Cnv_Settings : "Inbound_Cnv_Settings";
   END_VAR
   VAR_IN_OUT
      Cnv_Control : "Inbound_Cnv_Control_UDT";
      SinaSpeed : SinaSpeed;
   END_VAR
   VAR
      State : UInt;
      Timer_TC : TON_TIME;
      Timer_Transfer { S7_SetPoint := 'True'} : TON_TIME;
      Watchdog { S7_SetPoint := 'True'} : TON_TIME;
      Transfer_Direction { S7_SetPoint := 'True'} : String;
      MainSetpoint : Int;
      IEC_Timer_0_Instance_1 { S7_SetPoint := 'True'} : TON_TIME;
      R_TRIG_Instance { S7_SetPoint := 'True'} : R_TRIG;
   END_VAR
   VAR_TEMP
      Execute_Old : Bool;
      Stop_Old : Bool;
   END_VAR
BEGIN
   "R_TRIG_DB_8"(CLK:= #Cnv_Control.Instruction.Execute AND NOT #Execute_Old);
   "R_TRIG_DB_9"(CLK:=#Cnv_Control.Instruction.Stop AND NOT #Stop_Old);

   // "Debug_Barcode" := TRUE;

   #Execute_Old := #Cnv_Control.Instruction.Execute;
   #Stop_Old := #Cnv_Control.Instruction.Stop;

   #Cnv_Control.Enabled := #Cnv_Control.Instruction.Enable;

   //MODES
   #Cnv_Control.Mode := #Cnv_Control.Instruction.Mode_Change;
   IF (#Cnv_Control.Mode = 1 OR #Cnv_Control.Mode = 5) AND NOT #Cnv_Control.Error THEN
       #State := 500;
   END_IF;

   #R_TRIG_Instance(CLK:=#Cnv_Control.Mode = 3);
   IF #R_TRIG_Instance.Q THEN
       #State := 0;
   END_IF;

   (*
   TODO:
   01. Need to add statemachine watchdog - Done
   02. Extractor needs to be on same floor for pallet to be moved in manual passed Rbwd - Done
   03. Complete reset state - Done
   04. Add stop inputs - Done
   05. Need to add variable motor speed, manual needs to be slower. - Done
   06. Need to add cyclic error checking. For odd sensor combinations as well - Partially done
   07. Need to add Shuttle monitor - Done
   08. Need to add Task ID check and start bit check to outbound pallet move. Check direction of pallet movement based on connected Cnv.
   09. Need to add checks for wrong direction of travel - Done
   10. Add checks for unsafe conditions with Cnv_Inputs - Partially Done
   11. Define Error codes - DOne
   12. Add watchdof time to Cnv Settings - Done
   13. Add self-timeout on manual 
   14. For shuttle in place sensor checks take into account extractor floor and safety stopper state
   15. Confirm modes and states are correct (Semi-auto and maintenance as well)
   16. Add the correct transfer process for the logistex-spacemaker pallet handovers.

   Mode select is done via the HMI. Might add external mode select switches.

           Mode select mask:
           0: Disabled
           1: Manual
           2: Semi-Auto
           3: Auto
           4: Teach - N/A for Cnv
           5: Maintenance

   Device ID Format: XXYYZZ    
   XX = Device type   
       01   VTD
       10  Cnv_Front_of_VTD
       11  Cnv_Rear_of_VTD
       12  Cnv_On_Extractor
       20  Safety_Stop_Front_of_VTD
       21  Safety_Stop_Rear_of_VTD
   YY = Floor   
   ZZ = VTD Connected to    
   Example: 110203 Conveyor at the rear of VTD 3 on level 2

   Pallet Alignment
   0 = no alignment
   1 = center alignment
   2 = Left
   3 = Right

    Sensor order for the conveyor:
    Lfwd Lpd1 Lpd2
     []   []   []
    ##############################
    #        Pallet Flow         #
    #         ------->>          #
    #                            #
    #                            #
    ##############################
                     []   []   []
                    Rpd2 Rpd1 Rbwd      
   *)

   REGION Cyclic Checks    
       // Update the pallet type as the Cnv_Inputs are triggered.
       #Cnv_Control.Cnv_Occupied := NOT "Inbound Conveyor - Back Sensor" OR NOT "Inbound Conveyor - Front Sensor";

       // Update the Cnv_Control opbject
       #Cnv_Control.SM_State := #State;
       #Cnv_Control.Stopped := NOT #Cnv_Control.Running;
       IF #Cnv_Control.Instruction.Inbound_Ready OR #Cnv_Control.Instruction.Outbound_Ready THEN
           #Cnv_Control.Ready_For_Task := TRUE;
       ELSE
           #Cnv_Control.Ready_For_Task := FALSE;
       END_IF;

       //Automatic Start
       "IEC_Timer_0_DB_14".TON(IN := NOT #Cnv_Control.Inputs."Fork Lift Detect" AND #Cnv_Control.Inputs."Pallet Detect 1",
                               PT := UINT_TO_TIME(#Cnv_Settings.No_Forklift_Detect_Timer) * 1000);

       "IEC_Timer_0_DB_13".TP(IN:=#Cnv_Control.Inputs."Pallet Detect 1" AND "IEC_Timer_0_DB_14".Q,
                               PT:=T#3S,
                               Q=>#Cnv_Control.Instruction.Automatic_Start);

   END_REGION

   REGION Auto/Semi/Manual mode
       CASE #State OF
           0: //Initialization
               #Cnv_Control.Instruction.Transfer_Complete := 0;
               #Cnv_Control.Instruction.Transfer_in_Progress := FALSE;
               #Cnv_Control.Running := FALSE;
               #Cnv_Control.Motor.Forward := FALSE;
               #Cnv_Control.Motor.Reverse := FALSE;
               #Cnv_Control.Motor.Speed := 0;
               #Timer_Transfer(IN := FALSE,
                               PT := T#0S);
               IF #Cnv_Control.Enabled AND (#Cnv_Control.Mode = 3 OR #Cnv_Control.Mode = 2) AND #Cnv_Control.Error = 0 THEN
                   #State := 10;
               END_IF;

           10: // Idle - Waiting for Execute
               IF "R_TRIG_DB_8".Q AND NOT #Cnv_Control.Error THEN
                   #Cnv_Control.Done := FALSE;
                   #Cnv_Control.Running := TRUE;
                   #Cnv_Control.Motor.Forward := TRUE;
                   #Cnv_Control.Motor.Speed := #Cnv_Settings.Full_Speed;
                   #Transfer_Direction := 'Foward';
                   #Cnv_Control.Instruction.Transfer_in_Progress := TRUE;
                   #State := 20;//Without bacode
               ELSIF #Cnv_Control.Instruction.Start_Transfer AND NOT #Cnv_Control.Error AND
                   NOT "Inbound Conveyor - Back Sensor" AND "Inbound Conveyor - Front Sensor" THEN
                   #Cnv_Control.Done := FALSE;
                   #Cnv_Control.Running := TRUE;
                   #Cnv_Control.Motor.Forward := TRUE;
                   #Cnv_Control.Motor.Speed := #Cnv_Settings.Full_Speed;
                   #Transfer_Direction := 'Foward';
                   #Cnv_Control.Instruction.Transfer_in_Progress := TRUE;
                   #State := 15;
               END_IF;

           15: // Running Roller till the second sensor
               IF NOT "Inbound Conveyor - Front Sensor" THEN
                   #Cnv_Control.Motor.Speed := 0;
                   #Cnv_Control.Motor.Forward := FALSE;
                   #Cnv_Control.Running := FALSE;
                   #State := 20;
               END_IF;

               //Monitor the transfer progress
               #Timer_Transfer(IN := TRUE,
                               PT := UINT_TO_TIME(#Cnv_Settings.Transfer_Time) * 1000);
               //If the watchdog bites, kill the process
               IF #Timer_Transfer.Q THEN //14:1 Transfer timed out
                   "Set_Bit_F"(Bit := 3,
                               Bit_Value := 1,
                               Var := #Cnv_Control.Cnv_Errors.Error_Word_2);
               END_IF;


           20: //Read Barcode
               "IEC_Timer_0_DB_20".TON(IN:=TRUE,
                                       PT:=T#1S);

               IF "IEC_Timer_0_DB_20".Q OR "Control_DB".InBarcode_Station.Valid OR "Debug_Barcode" THEN
                   #State := 30;
               END_IF;

           30: //Wait PopUp 1 to run
               IF "Control_DB".PopUp_Cnv[1].Roller_Motor.Status.%X0 THEN
                   #Cnv_Control.Running := TRUE;
                   #Cnv_Control.Motor.Forward := TRUE;
                   #Cnv_Control.Motor.Speed := #Cnv_Settings.Full_Speed;
                   #Transfer_Direction := 'Foward';
                   #Cnv_Control.Instruction.Transfer_in_Progress := TRUE;
                   #State := 40;
               END_IF;

           40: // Running Roller
               IF "R_TRIG_DB_9".Q OR "PopUp Conveyor 2 - Pallet present 3" THEN
                   #Cnv_Control.Done := TRUE;
                   #Cnv_Control.Motor.Speed := 0;
                   #Cnv_Control.Motor.Forward := FALSE;
                   #Cnv_Control.Running := FALSE;
                   #State := 0;
               END_IF;

               //Monitor the transfer progress
               #Timer_Transfer(IN := TRUE,
                               PT := UINT_TO_TIME(#Cnv_Settings.Transfer_Time) * 1000);
               //If the watchdog bites, kill the process
               IF #Timer_Transfer.Q THEN //14:1 Transfer timed out
                   "Set_Bit_F"(Bit := 3,
                               Bit_Value := 1,
                               Var := #Cnv_Control.Cnv_Errors.Error_Word_2);
               END_IF;

               400: //Error state
                   #Cnv_Control.Running := FALSE;
                   #Cnv_Control.Motor.Speed := 0;
                   #Cnv_Control.Motor.Forward := FALSE;
                   #Cnv_Control.Motor.Reverse := FALSE;
                   #Cnv_Control.Instruction.Stop := FALSE;
                   #Cnv_Control.Instruction.Transfer_in_Progress := FALSE;
                   #Watchdog(IN := FALSE,
                                   PT := T#0S);
                   #Timer_TC(IN := FALSE,
                                   PT := T#0S);
                   #Timer_Transfer(IN := FALSE,
                                   PT := T#0S);
                   #IEC_Timer_0_Instance_1(IN := FALSE,
                                           PT := T#0S);
                   IF #Cnv_Control.Instruction.Reset THEN
                       #Cnv_Control.Warning := 0;
                       #Cnv_Control.Current_Task_ID := 0;
                       #Cnv_Control.Error := FALSE; //Reset the conveyor

                       #Cnv_Control.Cnv_Errors.Error_Word_1 := 0;
                       #Cnv_Control.Cnv_Errors.Error_Word_2 := 0;
                       #Cnv_Control.Cnv_Errors.Error_Word_3 := 0;
                       #Cnv_Control.Cnv_Errors.Error_Word_4 := 0;
                       #State := 0;
                   END_IF;

               500: //MANUAL MODE
                   IF #Cnv_Control.Enabled THEN
                       IF #Cnv_Control.Instruction.Foward OR #Cnv_Control.Instruction.Start_Transfer THEN
                           #Cnv_Control.Motor.Speed := #Cnv_Settings.Manual_Speed;
                           #Cnv_Control.Motor.Forward := TRUE;
                           #Cnv_Control.Running := TRUE;
                       ELSIF (#Cnv_Control.Instruction.Backward OR #Cnv_Control.Instruction.Start_Transfer_Backward) AND NOT #Cnv_Control.Inputs."Pallet Detect 1" THEN
                           #Cnv_Control.Motor.Speed := #Cnv_Settings.Manual_Speed;
                           #Cnv_Control.Motor.Reverse := TRUE;
                           #Cnv_Control.Running := TRUE;
                       ELSE
                           #Cnv_Control.Motor.Speed := 0;
                           #Cnv_Control.Motor.Forward := FALSE;
                           #Cnv_Control.Motor.Reverse := FALSE;
                           #Cnv_Control.Running := FALSE;
                       END_IF;
                   END_IF;
                   IF #Cnv_Control.Mode <> 1 AND #Cnv_Control.Mode <> 5 THEN
                       #State := 0;
                   END_IF;
           END_CASE;
       END_REGION



   REGION Cyclic Error Checks
       IF NOT "Main_Safety_RTG1_DB".SAFETY_OK_CAROUSEL THEN //11:1
           "Set_Bit_F"(Bit := 0,
                       Bit_Value := 1,
                       Var := #Cnv_Control.Cnv_Errors.Error_Word_1);
       END_IF;

       // IF #Cnv_Control.Instruction.Stop THEN //11:2
       //     "Set_Bit_F"(Bit := 1,
       //                 Bit_Value := 1,
       //                 Var := #Cnv_Control.Cnv_Errors.Error_Word_1);
       // END_IF;

       IF #Cnv_Control.Motor.Error THEN
           "Set_Bit_F"(Bit := 0,
                       Bit_Value := 1,
                       Var := #Cnv_Control.Cnv_Errors.Error_Word_4);
       END_IF;

       // Pallet Sensor Checks
       // IF #Cnv_Control.Inputs.Lfwd AND #Cnv_Control.Inputs.Rbwd THEN
       //     #Cnv_Control.Error := TRUE; //15:2 Combination of Cnv_Inputs indicates issue in conveyor
       //     "Set_Bit_F"(Bit := 1,
       //                 Bit_Value := 1,
       //                 Var := #Cnv_Control.Cnv_Errors.Error_Word_4);
       //     #State := 400;
       // IF #Cnv_Control.Inputs.Lfwd AND #Cnv_Control.Inputs.Lpd1 AND #Cnv_Control.Inputs.Rpd1 THEN
       //     #Cnv_Control.Error := TRUE; //15:3 Combination of Cnv_Inputs indicates issue in conveyor
       //     "Set_Bit_F"(Bit := 2,
       //                 Bit_Value := 1,
       //                 Var := #Cnv_Control.Cnv_Errors.Error_Word_4);
       //     #State := 400;
       // ELSIF #Cnv_Control.Inputs.Rbwd AND #Cnv_Control.Inputs.Lpd1 AND #Cnv_Control.Inputs.Rpd1 THEN
       //     #Cnv_Control.Error := TRUE; //15:4 Combination of Cnv_Inputs indicates issue in conveyor
       //     "Set_Bit_F"(Bit := 3,
       //                 Bit_Value := 1,
       //                 Var := #Cnv_Control.Cnv_Errors.Error_Word_4);
       //     #State := 400;
       // END_IF;

       // Shuttle in Place Cnv_Inputs - Need to confirm the order of these Cnv_Inputs.
       // IF (#Cnv_Settings.ID > 110000 AND #Cnv_Settings.ID < 120000 AND NOT #Cnv_Control.Inputs.Sdetect1 AND #Cnv_Control.Inputs.Sdetect2)
       //     OR (#Cnv_Settings.ID > 120000 AND #Cnv_Settings.ID < 130000 AND NOT #Cnv_Control.Inputs.Sdetect1 AND #Cnv_Control.Inputs.Sdetect2) THEN
       //     #Cnv_Control.Error := TRUE; //14:5 Shuttle is about to yeet itself down the VTD shaft
       //     "Set_Bit_F"(Bit := 7,
       //                 Bit_Value := 1,
       //                 Var := #Cnv_Control.Cnv_Errors.Error_Word_2);
       //     #State := 400;
       // END_IF;

       // IF (#Cnv_Settings.ID > 110000 AND #Cnv_Settings.ID < 120000 AND #Cnv_Control.Inputs.Sdetect1 AND NOT #Cnv_Control.Inputs.Sdetect2)
       //     OR (#Cnv_Settings.ID > 120000 AND #Cnv_Settings.ID < 130000 AND #Cnv_Control.Inputs.Sdetect1 AND NOT #Cnv_Control.Inputs.Sdetect2) THEN
       //     #Cnv_Control.Warning := 0; //Shuttle detected in conveyor not yet on barcode
       // END_IF;

       // // #Watchdog auto starts the moment Any form OF transfer occurs.
       // IF #State > 10 AND #State < 400 THEN
       //     #Watchdog(IN := TRUE,
       //               PT := T#200s);
       // ELSE
       //     #Watchdog.IN := FALSE;
       // END_IF;

       // IF #Watchdog.Q THEN
       //     #Watchdog.IN := FALSE;
       //     #Cnv_Control.Error := TRUE; //14:2  Watchdog bit
       //     "Set_Bit_F"(Bit := 4,
       //                 Bit_Value := 1,
       //                 Var := #Cnv_Control.Cnv_Errors.Error_Word_2);
       //     #State := 400;
       // END_IF;

       // go to error state
       IF #Cnv_Control.Cnv_Errors.Error_Word_1 <> 0 OR
           #Cnv_Control.Cnv_Errors.Error_Word_2 <> 0 OR
           #Cnv_Control.Cnv_Errors.Error_Word_3 <> 0 OR
           #Cnv_Control.Cnv_Errors.Error_Word_4 <> 0
           THEN
               #Cnv_Control.Error := TRUE;
               #State := 400;
       END_IF;
   END_REGION

   REGION VFD
       //Status
       #Cnv_Control.Motor.Ready := NOT #Cnv_Control.Motor.Error;

       #SinaSpeed(EnableAxis := #Cnv_Control.Motor.Forward OR #Cnv_Control.Motor.Reverse,
                  AckError := #Cnv_Control.Instruction.Reset,
                  SpeedSp := #MainSetpoint,
                  RefSpeed := 1745.0,
                  HWIDSTW := #Cnv_Settings.G120_Hardware_ID,
                  HWIDZSW := #Cnv_Settings.G120_Hardware_ID,
                  AxisEnabled => #Cnv_Control.Motor.Status.%X0,
                  Lockout => #Cnv_Control.Motor.Error,
                  Error => #Cnv_Control.Motor.Error);

       //MAIN SETPOINT
       IF #Cnv_Control.Motor.Forward THEN
           #MainSetpoint := (SCALE_X(MIN := 0,
                                    VALUE := NORM_X(MIN := 0,
                                                    VALUE := #Cnv_Control.Motor.Speed,
                                                    MAX := 100),
                                    MAX := 1745.0) * -1);
       ELSIF #Cnv_Control.Motor.Reverse THEN
           #MainSetpoint := SCALE_X(MIN := 0,
                                     VALUE := NORM_X(MIN := 0,
                                                     VALUE := #Cnv_Control.Motor.Speed,
                                                     MAX := 100),
                                     MAX := 1745.0);
       ELSE
           #MainSetpoint := 0;
       END_IF;


       REGION Actual Speed
           IF #MainSetpoint > 0 THEN
               #Cnv_Control.Motor.Speed_Actual := SCALE_X(MIN := 0,
                                                          VALUE := NORM_X(MIN := 0,
                                                                          VALUE := #SinaSpeed.ActVelocity,
                                                                          MAX := 1745.0),
                                                          MAX := 100);
           ELSIF #MainSetpoint < 0 THEN
               #Cnv_Control.Motor.Speed_Actual := SCALE_X(MIN := 0,
                                                          VALUE := NORM_X(MIN := 0,
                                                                          VALUE := #SinaSpeed.ActVelocity * -1,
                                                                          MAX := 1745.0),
                                                          MAX := 100);
           ELSE
               #Cnv_Control.Motor.Speed_Actual := 0;
           END_IF;
       END_REGION
   END_REGION
END_FUNCTION_BLOCK

FUNCTION_BLOCK "OutConveyor_FB"   // FB16, SCL
TITLE = Conveyor Instance FB
{ S7_Optimized_Access := 'TRUE' }
AUTHOR : Mertin Coetzee
VERSION : 0.1
// stored: AutoNumber true, IsIECCheckEnabled false, IsRetainMemResEnabled false, MemoryReserve 100, SetENOAutomatically false, UDAEnableTagReadback false
   VAR_INPUT
      Cnv_Settings : "Outbound_Cnv_Settings";
   END_VAR
   VAR_IN_OUT
      Cnv_Control : "Outbound_Cnv_Control";
      SinaSpeed : SinaSpeed;
   END_VAR
   VAR
      State : UInt;
      Timer_TC : TON_TIME;
      Timer_Transfer { S7_SetPoint := 'True'} : TON_TIME;
      Watchdog { S7_SetPoint := 'True'} : TON_TIME;
      Transfer_Direction { S7_SetPoint := 'True'} : String;
      MainSetpoint : Int;
      IEC_Timer_0_Instance_1 { S7_SetPoint := 'True'} : TON_TIME;
      R_TRIG_Instance { S7_SetPoint := 'True'} : R_TRIG;
   END_VAR
   VAR_TEMP
      Execute_Old : Bool;
      Stop_Old : Bool;
   END_VAR
BEGIN
   "R_TRIG_DB_11"(CLK := #Cnv_Control.Instruction.Execute AND NOT #Execute_Old);
   "R_TRIG_DB_12"(CLK := #Cnv_Control.Instruction.Stop AND NOT #Stop_Old);

   #Execute_Old := #Cnv_Control.Instruction.Execute;
   #Stop_Old := #Cnv_Control.Instruction.Stop;

